// TIA Portal V20 program export: 15 tag tables, 7 data types, 9 data blocks, 10 code blocks (in call order from the OBs), 5 instance data blocks

VAR_GLOBAL   // PLC tag table "COGNEX_ETIKETA"
   "COG_ETIKETA_COG_ETIKETA_is3800-TriggerEnable" AT %Q2.0 : Bool;
   "COG_ETIKETA_COG_ETIKETA_is3800-Trigger" AT %Q2.1 : Bool;
   "COG_ETIKETA_is3800-ClearExposureComplete" AT %Q2.2 : Bool;
   "COG_ETIKETA_is3800-Set Offline" AT %Q2.7 : Bool;
   "COG_ETIKETA_is3800-TriggerReady" AT %I2.0 : Bool;
   "COG_ETIKETA_is3800-TriggerAck" AT %I2.1 : Bool;
   "COG_ETIKETA_is3800-ExposureComplete" AT %I2.2 : Bool;
   "COG_ETIKETA_is3800-AcquCOG_ETIKETA_isitionError" AT %I2.3 : Bool;
   "COG_ETIKETA_is3800-Offline Reason" AT %I2.4 : Bool;
   "COG_ETIKETA_is3800-Offline Reason(1)" AT %I2.5 : Bool;
   "COG_ETIKETA_is3800-Offline Reason(2)" AT %I2.6 : Bool;
   "COG_ETIKETA_is3800-Online" AT %I2.7 : Bool;
   "COG_ETIKETA_is3800-AcquCOG_ETIKETA_isitionID" AT %IW4 : Int;
   "COG_ETIKETA_is3800-BufferResultsEnable" AT %Q3.0 : Bool;
   "COG_ETIKETA_is3800-InspectionResultsAck" AT %Q3.1 : Bool;
   "COG_ETIKETA_is3800-SetUserData" AT %Q3.2 : Bool;
   "COG_ETIKETA_is3800-ExecuteCommand/JobLoad" AT %Q3.3 : Bool;
   "COG_ETIKETA_is3800-ClearError" AT %Q3.7 : Bool;
   "COG_ETIKETA_is3800-Reserved" AT %I10.0 : Bool;
   "COG_ETIKETA_is3800-InspectionCompleted" AT %I10.1 : Bool;
   "COG_ETIKETA_is3800-ResultsBufferOverrun" AT %I10.2 : Bool;
   "COG_ETIKETA_is3800-ResultsValid" AT %I10.3 : Bool;
   "COG_ETIKETA_is3800-CommandExecuting" AT %I10.4 : Bool;
   "COG_ETIKETA_is3800-CommandCompleted" AT %I10.5 : Bool;
   "COG_ETIKETA_is3800-CommandFailed" AT %I10.6 : Bool;
   "COG_ETIKETA_is3800-SetUserDataAck" AT %I10.7 : Bool;
   "COG_ETIKETA_is3800-ResultsPassed (Job)" AT %I11.0 : Bool;
   "COG_ETIKETA_is3800-SystemValidated" AT %I11.1 : Bool;
   "COG_ETIKETA_is3800-Error" AT %I11.7 : Bool;
   "COG_ETIKETA_is3800-ErrorCode" AT %IW12 : Word;
   "COG_ETIKETA_is3800-CommandID" AT %QW64 : Word;
   "COG_ETIKETA_is3800-Current Job ID" AT %IW68 : Word;
   "COG_ETIKETA_is3800-CommandResultCode" AT %IW70 : Word;
   "COG_ETIKETA_is3800-ExternalEvent[0]" AT %Q4.0 : Bool;
   "COG_ETIKETA_is3800-ExternalEvent[1]" AT %Q4.1 : Bool;
   "COG_ETIKETA_is3800-ExternalEvent[2]" AT %Q4.2 : Bool;
   "COG_ETIKETA_is3800-ExternalEvent[3]" AT %Q4.3 : Bool;
   "COG_ETIKETA_is3800-ExternalEvent[4]" AT %Q4.4 : Bool;
   "COG_ETIKETA_is3800-ExternalEvent[5]" AT %Q4.5 : Bool;
   "COG_ETIKETA_is3800-ExternalEvent[6]" AT %Q4.6 : Bool;
   "COG_ETIKETA_is3800-ExternalEvent[7]" AT %Q4.7 : Bool;
   "COG_ETIKETA_is3800-ExternalEventAck[0]" AT %I6.0 : Bool;
   "COG_ETIKETA_is3800-ExternalEventAck[1]" AT %I6.1 : Bool;
   "COG_ETIKETA_is3800-ExternalEventAck[2]" AT %I6.2 : Bool;
   "COG_ETIKETA_is3800-ExternalEventAck[3]" AT %I6.3 : Bool;
   "COG_ETIKETA_is3800-ExternalEventAck[4]" AT %I6.4 : Bool;
   "COG_ETIKETA_is3800-ExternalEventAck[5]" AT %I6.5 : Bool;
   "COG_ETIKETA_is3800-ExternalEventAck[6]" AT %I6.6 : Bool;
   "COG_ETIKETA_is3800-ExternalEventAck[7]" AT %I6.7 : Bool;
   "COG_ETIKETA_is3800-UserData[0]" AT %QB66 : Byte;
   "COG_ETIKETA_is3800-UserData[1]" AT %QB67 : Byte;
   "COG_ETIKETA_is3800-UserData[2]" AT %QB68 : Byte;
   "COG_ETIKETA_is3800-UserData[3]" AT %QB69 : Byte;
   "COG_ETIKETA_is3800-UserData[4]" AT %QB70 : Byte;
   "COG_ETIKETA_is3800-UserData[5]" AT %QB71 : Byte;
   "COG_ETIKETA_is3800-UserData[6]" AT %QB72 : Byte;
   "COG_ETIKETA_is3800-UserData[7]" AT %QB73 : Byte;
   "COG_ETIKETA_is3800-UserData[8]" AT %QB74 : Byte;
   "COG_ETIKETA_is3800-UserData[9]" AT %QB75 : Byte;
   "COG_ETIKETA_is3800-UserData[10]" AT %QB76 : Byte;
   "COG_ETIKETA_is3800-UserData[11]" AT %QB77 : Byte;
   "COG_ETIKETA_is3800-UserData[12]" AT %QB78 : Byte;
   "COG_ETIKETA_is3800-UserData[13]" AT %QB79 : Byte;
   "COG_ETIKETA_is3800-UserData[14]" AT %QB80 : Byte;
   "COG_ETIKETA_is3800-UserData[15]" AT %QB81 : Byte;
   "COG_ETIKETA_is3800-InspectionID" AT %IW72 : Word;
   "COG_ETIKETA_is3800-InspectionResultsCode" AT %IW74 : Int;
   "COG_ETIKETA_is3800-InspectionResults_0" AT %IB76 : Byte;
   "COG_ETIKETA_is3800-InspectionResults_1" AT %IB77 : Byte;
   "COG_ETIKETA_is3800-InspectionResults_2" AT %IB78 : Byte;
   "COG_ETIKETA_is3800-InspectionResults_3" AT %IB79 : Byte;
   "COG_ETIKETA_is3800-InspectionResults_4" AT %IB80 : Byte;
   "COG_ETIKETA_is3800-InspectionResults_5" AT %IB81 : Byte;
   "COG_ETIKETA_is3800-InspectionResults_6" AT %IB82 : Byte;
   "COG_ETIKETA_is3800-InspectionResults_7" AT %IB83 : Byte;
   "COG_ETIKETA_is3800-InspectionResults_8" AT %IB84 : Byte;
   "COG_ETIKETA_is3800-InspectionResults_9" AT %IB85 : Byte;
   "COG_ETIKETA_is3800-InspectionResults_10" AT %IB86 : Byte;
   "COG_ETIKETA_is3800-InspectionResults_11" AT %IB87 : Byte;
   "COG_ETIKETA_is3800-InspectionResults_12" AT %IB88 : Byte;
   "COG_ETIKETA_is3800-InspectionResults_13" AT %IB89 : Byte;
   "COG_ETIKETA_is3800-InspectionResults_14" AT %IB90 : Byte;
   "COG_ETIKETA_is3800-InspectionResults_15" AT %IB91 : Byte;
   "COG_ETIKETA_is3800-InspectionResults_16" AT %IB92 : Byte;
   "COG_ETIKETA_is3800-InspectionResults_17" AT %IB93 : Byte;
   "COG_ETIKETA_is3800-InspectionResults_18" AT %IB94 : Byte;
   "COG_ETIKETA_is3800-InspectionResults_19" AT %IB95 : Byte;
   "COG_ETIKETA_is3800-InspectionResults_20" AT %IB96 : Byte;
   "COG_ETIKETA_is3800-InspectionResults_21" AT %IB97 : Byte;
   "COG_ETIKETA_is3800-InspectionResults_22" AT %IB98 : Byte;
   "COG_ETIKETA_is3800-InspectionResults_23" AT %IB99 : Byte;
   "COG_ETIKETA_is3800-InspectionResults_24" AT %IB100 : Byte;
   "COG_ETIKETA_is3800-InspectionResults_25" AT %IB101 : Byte;
   "COG_ETIKETA_is3800-InspectionResults_26" AT %IB102 : Byte;
   "COG_ETIKETA_is3800-InspectionResults_27" AT %IB103 : Byte;
   "COG_ETIKETA_is3800-InspectionResults_28" AT %IB104 : Byte;
   "COG_ETIKETA_is3800-InspectionResults_29" AT %IB105 : Byte;
   "COG_ETIKETA_is3800-InspectionResults_30" AT %IB106 : Byte;
   "COG_ETIKETA_is3800-InspectionResults_31" AT %IB107 : Byte;
   "COG_ETIKETA_is3800-InspectionResults_32" AT %IB108 : Byte;
   "COG_ETIKETA_is3800-InspectionResults_33" AT %IB109 : Byte;
   "COG_ETIKETA_is3800-InspectionResults_34" AT %IB110 : Byte;
   "COG_ETIKETA_is3800-InspectionResults_35" AT %IB111 : Byte;
   "COG_ETIKETA_is3800-InspectionResults_36" AT %IB112 : Byte;
   "COG_ETIKETA_is3800-InspectionResults_37" AT %IB113 : Byte;
   "COG_ETIKETA_is3800-InspectionResults_38" AT %IB114 : Byte;
   "COG_ETIKETA_is3800-InspectionResults_39" AT %IB115 : Byte;
   "COG_ETIKETA_is3800-InspectionResults_40" AT %IB116 : Byte;
   "COG_ETIKETA_is3800-InspectionResults_41" AT %IB117 : Byte;
   "COG_ETIKETA_is3800-InspectionResults_42" AT %IB118 : Byte;
   "COG_ETIKETA_is3800-InspectionResults_43" AT %IB119 : Byte;
   "COG_ETIKETA_is3800-InspectionResults_44" AT %IB120 : Byte;
   "COG_ETIKETA_is3800-InspectionResults_45" AT %IB121 : Byte;
   "COG_ETIKETA_is3800-InspectionResults_46" AT %IB122 : Byte;
   "COG_ETIKETA_is3800-InspectionResults_47" AT %IB123 : Byte;
   "COG_ETIKETA_is3800-InspectionResults_48" AT %IB124 : Byte;
   "COG_ETIKETA_is3800-InspectionResults_49" AT %IB125 : Byte;
   "COG_ETIKETA_is3800-InspectionResults_50" AT %IB126 : Byte;
   "COG_ETIKETA_is3800-InspectionResults_51" AT %IB127 : Byte;
   "COG_ETIKETA_is3800-InspectionResults_52" AT %IB128 : Byte;
   "COG_ETIKETA_is3800-InspectionResults_53" AT %IB129 : Byte;
   "COG_ETIKETA_is3800-InspectionResults_54" AT %IB130 : Byte;
   "COG_ETIKETA_is3800-InspectionResults_55" AT %IB131 : Byte;
   "COG_ETIKETA_is3800-InspectionResults_56" AT %IB132 : Byte;
   "COG_ETIKETA_is3800-InspectionResults_57" AT %IB133 : Byte;
   "COG_ETIKETA_is3800-InspectionResults_58" AT %IB134 : Byte;
   "COG_ETIKETA_is3800-InspectionResults_59" AT %IB135 : Byte;
   "COG_ETIKETA_is3800-InspectionResults_60" AT %IB136 : Byte;
   "COG_ETIKETA_is3800-InspectionResults_61" AT %IB137 : Byte;
   "COG_ETIKETA_is3800-InspectionResults_62" AT %IB138 : Byte;
   "COG_ETIKETA_is3800-InspectionResults_63" AT %IB139 : Byte;
   "COG_ETIKETA_is3800-InspectionResults_64" AT %IB140 : Byte;
   "COG_ETIKETA_is3800-InspectionResults_65" AT %IB141 : Byte;
   "COG_ETIKETA_is3800-InspectionResults_66" AT %IB142 : Byte;
   "COG_ETIKETA_is3800-InspectionResults_67" AT %IB143 : Byte;
   "COG_ETIKETA_is3800-InspectionResults_68" AT %IB144 : Byte;
   "COG_ETIKETA_is3800-InspectionResults_69" AT %IB145 : Byte;
   "COG_ETIKETA_is3800-InspectionResults_70" AT %IB146 : Byte;
   "COG_ETIKETA_is3800-InspectionResults_71" AT %IB147 : Byte;
   "COG_ETIKETA_is3800-InspectionResults_72" AT %IB148 : Byte;
   "COG_ETIKETA_is3800-InspectionResults_73" AT %IB149 : Byte;
   "COG_ETIKETA_is3800-InspectionResults_74" AT %IB150 : Byte;
   "COG_ETIKETA_is3800-InspectionResults_75" AT %IB151 : Byte;
   "COG_ETIKETA_is3800-InspectionResults_76" AT %IB152 : Byte;
   "COG_ETIKETA_is3800-InspectionResults_77" AT %IB153 : Byte;
   "COG_ETIKETA_is3800-InspectionResults_78" AT %IB154 : Byte;
   "COG_ETIKETA_is3800-InspectionResults_79" AT %IB155 : Byte;
   "COG_ETIKETA_is3800-InspectionResults_80" AT %IB156 : Byte;
   "COG_ETIKETA_is3800-InspectionResults_81" AT %IB157 : Byte;
   "COG_ETIKETA_is3800-InspectionResults_82" AT %IB158 : Byte;
   "COG_ETIKETA_is3800-InspectionResults_83" AT %IB159 : Byte;
   "COG_ETIKETA_is3800-InspectionResults_84" AT %IB160 : Byte;
   "COG_ETIKETA_is3800-InspectionResults_85" AT %IB164 : Byte;
   "COG_ETIKETA_is3800-InspectionResults_86" AT %IB165 : Byte;
   "COG_ETIKETA_is3800-InspectionResults_87" AT %IB166 : Byte;
   "COG_ETIKETA_is3800-InspectionResults_88" AT %IB167 : Byte;
   "COG_ETIKETA_is3800-InspectionResults_89" AT %IB168 : Byte;
   "COG_ETIKETA_is3800-InspectionResults_90" AT %IB169 : Byte;
   "COG_ETIKETA_is3800-InspectionResults_91" AT %IB170 : Byte;
   "COG_ETIKETA_is3800-InspectionResults_92" AT %IB171 : Byte;
   "COG_ETIKETA_is3800-InspectionResults_93" AT %IB172 : Byte;
   "COG_ETIKETA_is3800-InspectionResults_94" AT %IB173 : Byte;
   "COG_ETIKETA_is3800-InspectionResults_95" AT %IB174 : Byte;
   "COG_ETIKETA_is3800-InspectionResults_96" AT %IB175 : Byte;
   "COG_ETIKETA_is3800-InspectionResults_97" AT %IB176 : Byte;
   "COG_ETIKETA_is3800-InspectionResults_98" AT %IB177 : Byte;
   "COG_ETIKETA_is3800-InspectionResults_99" AT %IB178 : Byte;
   "COG_ETIKETA_is3800-InspectionResults_100" AT %IB179 : Byte;
END_VAR

VAR_GLOBAL   // PLC tag table "COGNEX_FOLIE_L"
   "COG_FOLIE_L_COG_FOLIE_L_is3800-TriggerEnable" AT %Q5.0 : Bool;
   "COG_FOLIE_L_is3800-Trigger" AT %Q5.1 : Bool;
   "COG_FOLIE_L_is3800-ClearExposureComplete" AT %Q5.2 : Bool;
   "COG_FOLIE_L_is3800-Set Offline" AT %Q5.7 : Bool;
   "COG_FOLIE_L_is3800-TriggerReady" AT %I14.0 : Bool;
   "COG_FOLIE_L_is3800-TriggerAck" AT %I14.1 : Bool;
   "COG_FOLIE_L_is3800-ExposureComplete" AT %I14.2 : Bool;
   "COG_FOLIE_L_is3800-AcquCOG_FOLIE_L_isitionError" AT %I14.3 : Bool;
   "COG_FOLIE_L_is3800-Offline Reason" AT %I14.4 : Bool;
   "COG_FOLIE_L_is3800-Offline Reason(1)" AT %I14.5 : Bool;
   "COG_FOLIE_L_is3800-Offline Reason(2)" AT %I14.6 : Bool;
   "COG_FOLIE_L_is3800-Online" AT %I14.7 : Bool;
   "COG_FOLIE_L_is3800-AcquCOG_FOLIE_L_isitionID" AT %IW16 : Int;
   "COG_FOLIE_L_is3800-BufferResultsEnable" AT %Q6.0 : Bool;
   "COG_FOLIE_L_is3800-InspectionResultsAck" AT %Q6.1 : Bool;
   "COG_FOLIE_L_is3800-SetUserData" AT %Q6.2 : Bool;
   "COG_FOLIE_L_is3800-ExecuteCommand/JobLoad" AT %Q6.3 : Bool;
   "COG_FOLIE_L_is3800-ClearError" AT %Q6.7 : Bool;
   "COG_FOLIE_L_is3800-Reserved" AT %I18.0 : Bool;
   "COG_FOLIE_L_is3800-InspectionCompleted" AT %I18.1 : Bool;
   "COG_FOLIE_L_is3800-ResultsBufferOverrun" AT %I18.2 : Bool;
   "COG_FOLIE_L_is3800-ResultsValid" AT %I18.3 : Bool;
   "COG_FOLIE_L_is3800-CommandExecuting" AT %I18.4 : Bool;
   "COG_FOLIE_L_is3800-CommandCompleted" AT %I18.5 : Bool;
   "COG_FOLIE_L_is3800-CommandFailed" AT %I18.6 : Bool;
   "COG_FOLIE_L_is3800-SetUserDataAck" AT %I18.7 : Bool;
   "COG_FOLIE_L_is3800-ResultsPassed (Job)" AT %I19.0 : Bool;
   "COG_FOLIE_L_is3800-SystemValidated" AT %I19.1 : Bool;
   "COG_FOLIE_L_is3800-Error" AT %I19.7 : Bool;
   "COG_FOLIE_L_is3800-ErrorCode" AT %IW20 : Word;
   "COG_FOLIE_L_is3800-CommandID" AT %QW130 : Word;
   "COG_FOLIE_L_is3800-Current Job ID" AT %IW140 : Word;
   "COG_FOLIE_L_is3800-CommandResultCode" AT %IW142 : Word;
   "COG_FOLIE_L_is3800-ExternalEvent[0]" AT %Q7.0 : Bool;
   "COG_FOLIE_L_is3800-ExternalEvent[1]" AT %Q7.1 : Bool;
   "COG_FOLIE_L_is3800-ExternalEvent[2]" AT %Q7.2 : Bool;
   "COG_FOLIE_L_is3800-ExternalEvent[3]" AT %Q7.3 : Bool;
   "COG_FOLIE_L_is3800-ExternalEvent[4]" AT %Q7.4 : Bool;
   "COG_FOLIE_L_is3800-ExternalEvent[5]" AT %Q7.5 : Bool;
   "COG_FOLIE_L_is3800-ExternalEvent[6]" AT %Q7.6 : Bool;
   "COG_FOLIE_L_is3800-ExternalEvent[7]" AT %Q7.7 : Bool;
   "COG_FOLIE_L_is3800-ExternalEventAck[0]" AT %I7.0 : Bool;
   "COG_FOLIE_L_is3800-ExternalEventAck[1]" AT %I7.1 : Bool;
   "COG_FOLIE_L_is3800-ExternalEventAck[2]" AT %I7.2 : Bool;
   "COG_FOLIE_L_is3800-ExternalEventAck[3]" AT %I7.3 : Bool;
   "COG_FOLIE_L_is3800-ExternalEventAck[4]" AT %I7.4 : Bool;
   "COG_FOLIE_L_is3800-ExternalEventAck[5]" AT %I7.5 : Bool;
   "COG_FOLIE_L_is3800-ExternalEventAck[6]" AT %I7.6 : Bool;
   "COG_FOLIE_L_is3800-ExternalEventAck[7]" AT %I7.7 : Bool;
   "COG_FOLIE_L_is3800-UserData[0]" AT %QB132 : Byte;
   "COG_FOLIE_L_is3800-UserData[1]" AT %QB133 : Byte;
   "COG_FOLIE_L_is3800-UserData[2]" AT %QB134 : Byte;
   "COG_FOLIE_L_is3800-UserData[3]" AT %QB135 : Byte;
   "COG_FOLIE_L_is3800-UserData[4]" AT %QB136 : Byte;
   "COG_FOLIE_L_is3800-UserData[5]" AT %QB137 : Byte;
   "COG_FOLIE_L_is3800-UserData[6]" AT %QB138 : Byte;
   "COG_FOLIE_L_is3800-UserData[7]" AT %QB139 : Byte;
   "COG_FOLIE_L_is3800-UserData[8]" AT %QB140 : Byte;
   "COG_FOLIE_L_is3800-UserData[9]" AT %QB141 : Byte;
   "COG_FOLIE_L_is3800-UserData[10]" AT %QB142 : Byte;
   "COG_FOLIE_L_is3800-UserData[11]" AT %QB143 : Byte;
   "COG_FOLIE_L_is3800-UserData[12]" AT %QB144 : Byte;
   "COG_FOLIE_L_is3800-UserData[13]" AT %QB145 : Byte;
   "COG_FOLIE_L_is3800-UserData[14]" AT %QB146 : Byte;
   "COG_FOLIE_L_is3800-UserData[15]" AT %QB147 : Byte;
   "COG_FOLIE_L_is3800-InspectionID" AT %IW144 : Word;
   "COG_FOLIE_L_is3800-InspectionResultsCode" AT %IW146 : Int;
   "COG_FOLIE_L_is3800-InspectionResults[0]" AT %IB148 : Byte;
   "COG_FOLIE_L_is3800-InspectionResults[1]" AT %IB149 : Byte;
   "COG_FOLIE_L_is3800-InspectionResults[2]" AT %IB150 : Byte;
   "COG_FOLIE_L_is3800-InspectionResults[3]" AT %IB151 : Byte;
   "COG_FOLIE_L_is3800-InspectionResults[4]" AT %IB152 : Byte;
   "COG_FOLIE_L_is3800-InspectionResults[5]" AT %IB153 : Byte;
   "COG_FOLIE_L_is3800-InspectionResults[6]" AT %IB154 : Byte;
   "COG_FOLIE_L_is3800-InspectionResults[7]" AT %IB155 : Byte;
   "COG_FOLIE_L_is3800-InspectionResults[8]" AT %IB156 : Byte;
   "COG_FOLIE_L_is3800-InspectionResults[9]" AT %IB157 : Byte;
   "COG_FOLIE_L_is3800-InspectionResults[10]" AT %IB158 : Byte;
   "COG_FOLIE_L_is3800-InspectionResults[11]" AT %IB159 : Byte;
   "COG_FOLIE_L_is3800-InspectionResults[12]" AT %IB160 : Byte;
   "COG_FOLIE_L_is3800-InspectionResults[13]" AT %IB161 : Byte;
   "COG_FOLIE_L_is3800-InspectionResults[14]" AT %IB162 : Byte;
   "COG_FOLIE_L_is3800-InspectionResults[15]" AT %IB163 : Byte;
END_VAR

VAR_GLOBAL   // PLC tag table "COGNEX_FOLIE_P"
   "COG_FOLIE_P_COG_FOLIE_P_is3800-TriggerEnable" AT %Q10.0 : Bool;
   "COG_FOLIE_P_is3800-Trigger" AT %Q10.1 : Bool;
   "COG_FOLIE_P_is3800-ClearExposureComplete" AT %Q10.2 : Bool;
   "COG_FOLIE_P_is3800-Set Offline" AT %Q10.7 : Bool;
   "COG_FOLIE_P_is3800-TriggerReady" AT %I22.0 : Bool;
   "COG_FOLIE_P_is3800-TriggerAck" AT %I22.1 : Bool;
   "COG_FOLIE_P_is3800-ExposureComplete" AT %I22.2 : Bool;
   "COG_FOLIE_P_is3800-AcquCOG_FOLIE_P_isitionError" AT %I22.3 : Bool;
   "COG_FOLIE_P_is3800-Offline Reason" AT %I22.4 : Bool;
   "COG_FOLIE_P_is3800-Offline Reason(1)" AT %I22.5 : Bool;
   "COG_FOLIE_P_is3800-Offline Reason(2)" AT %I22.6 : Bool;
   "COG_FOLIE_P_is3800-Online" AT %I22.7 : Bool;
   "COG_FOLIE_P_is3800-AcquCOG_FOLIE_P_isitionID" AT %IW24 : Int;
   "COG_FOLIE_P_is3800-BufferResultsEnable" AT %Q11.0 : Bool;
   "COG_FOLIE_P_is3800-InspectionResultsAck" AT %Q11.1 : Bool;
   "COG_FOLIE_P_is3800-SetUserData" AT %Q11.2 : Bool;
   "COG_FOLIE_P_is3800-ExecuteCommand/JobLoad" AT %Q11.3 : Bool;
   "COG_FOLIE_P_is3800-ClearError" AT %Q11.7 : Bool;
   "COG_FOLIE_P_is3800-Reserved" AT %I26.0 : Bool;
   "COG_FOLIE_P_is3800-InspectionCompleted" AT %I26.1 : Bool;
   "COG_FOLIE_P_is3800-ResultsBufferOverrun" AT %I26.2 : Bool;
   "COG_FOLIE_P_is3800-ResultsValid" AT %I26.3 : Bool;
   "COG_FOLIE_P_is3800-CommandExecuting" AT %I26.4 : Bool;
   "COG_FOLIE_P_is3800-CommandCompleted" AT %I26.5 : Bool;
   "COG_FOLIE_P_is3800-CommandFailed" AT %I26.6 : Bool;
   "COG_FOLIE_P_is3800-SetUserDataAck" AT %I26.7 : Bool;
   "COG_FOLIE_P_is3800-ResultsPassed (Job)" AT %I27.0 : Bool;
   "COG_FOLIE_P_is3800-SystemValidated" AT %I27.1 : Bool;
   "COG_FOLIE_P_is3800-Error" AT %I27.7 : Bool;
   "COG_FOLIE_P_is3800-ErrorCode" AT %IW28 : Word;
   "COG_FOLIE_P_is3800-CommandID" AT %QW196 : Word;
   "COG_FOLIE_P_is3800-Current Job ID" AT %IW212 : Word;
   "COG_FOLIE_P_is3800-CommandResultCode" AT %IW214 : Word;
   "COG_FOLIE_P_is3800-ExternalEvent[0]" AT %Q12.0 : Bool;
   "COG_FOLIE_P_is3800-ExternalEvent[1]" AT %Q12.1 : Bool;
   "COG_FOLIE_P_is3800-ExternalEvent[2]" AT %Q12.2 : Bool;
   "COG_FOLIE_P_is3800-ExternalEvent[3]" AT %Q12.3 : Bool;
   "COG_FOLIE_P_is3800-ExternalEvent[4]" AT %Q12.4 : Bool;
   "COG_FOLIE_P_is3800-ExternalEvent[5]" AT %Q12.5 : Bool;
   "COG_FOLIE_P_is3800-ExternalEvent[6]" AT %Q12.6 : Bool;
   "COG_FOLIE_P_is3800-ExternalEvent[7]" AT %Q12.7 : Bool;
   "COG_FOLIE_P_is3800-ExternalEventAck[0]" AT %I30.0 : Bool;
   "COG_FOLIE_P_is3800-ExternalEventAck[1]" AT %I30.1 : Bool;
   "COG_FOLIE_P_is3800-ExternalEventAck[2]" AT %I30.2 : Bool;
   "COG_FOLIE_P_is3800-ExternalEventAck[3]" AT %I30.3 : Bool;
   "COG_FOLIE_P_is3800-ExternalEventAck[4]" AT %I30.4 : Bool;
   "COG_FOLIE_P_is3800-ExternalEventAck[5]" AT %I30.5 : Bool;
   "COG_FOLIE_P_is3800-ExternalEventAck[6]" AT %I30.6 : Bool;
   "COG_FOLIE_P_is3800-ExternalEventAck[7]" AT %I30.7 : Bool;
   "COG_FOLIE_P_is3800-UserData[0]" AT %QB198 : Byte;
   "COG_FOLIE_P_is3800-UserData[1]" AT %QB199 : Byte;
   "COG_FOLIE_P_is3800-UserData[2]" AT %QB200 : Byte;
   "COG_FOLIE_P_is3800-UserData[3]" AT %QB201 : Byte;
   "COG_FOLIE_P_is3800-UserData[4]" AT %QB202 : Byte;
   "COG_FOLIE_P_is3800-UserData[5]" AT %QB203 : Byte;
   "COG_FOLIE_P_is3800-UserData[6]" AT %QB204 : Byte;
   "COG_FOLIE_P_is3800-UserData[7]" AT %QB205 : Byte;
   "COG_FOLIE_P_is3800-UserData[8]" AT %QB206 : Byte;
   "COG_FOLIE_P_is3800-UserData[9]" AT %QB207 : Byte;
   "COG_FOLIE_P_is3800-UserData[10]" AT %QB208 : Byte;
   "COG_FOLIE_P_is3800-UserData[11]" AT %QB209 : Byte;
   "COG_FOLIE_P_is3800-UserData[12]" AT %QB210 : Byte;
   "COG_FOLIE_P_is3800-UserData[13]" AT %QB211 : Byte;
   "COG_FOLIE_P_is3800-UserData[14]" AT %QB212 : Byte;
   "COG_FOLIE_P_is3800-UserData[15]" AT %QB213 : Byte;
   "COG_FOLIE_P_is3800-InspectionID" AT %IW216 : Word;
   "COG_FOLIE_P_is3800-InspectionResultsCode" AT %IW218 : Int;
   "COG_FOLIE_P_is3800-InspectionResults[0]" AT %IB220 : Byte;
   "COG_FOLIE_P_is3800-InspectionResults[1]" AT %IB221 : Byte;
   "COG_FOLIE_P_is3800-InspectionResults[2]" AT %IB222 : Byte;
   "COG_FOLIE_P_is3800-InspectionResults[3]" AT %IB223 : Byte;
   "COG_FOLIE_P_is3800-InspectionResults[4]" AT %IB224 : Byte;
   "COG_FOLIE_P_is3800-InspectionResults[5]" AT %IB225 : Byte;
   "COG_FOLIE_P_is3800-InspectionResults[6]" AT %IB226 : Byte;
   "COG_FOLIE_P_is3800-InspectionResults[7]" AT %IB227 : Byte;
   "COG_FOLIE_P_is3800-InspectionResults[8]" AT %IB228 : Byte;
   "COG_FOLIE_P_is3800-InspectionResults[9]" AT %IB229 : Byte;
   "COG_FOLIE_P_is3800-InspectionResults[10]" AT %IB230 : Byte;
   "COG_FOLIE_P_is3800-InspectionResults[11]" AT %IB231 : Byte;
   "COG_FOLIE_P_is3800-InspectionResults[12]" AT %IB232 : Byte;
   "COG_FOLIE_P_is3800-InspectionResults[13]" AT %IB233 : Byte;
   "COG_FOLIE_P_is3800-InspectionResults[14]" AT %IB234 : Byte;
   "COG_FOLIE_P_is3800-InspectionResults[15]" AT %IB235 : Byte;
END_VAR

VAR_GLOBAL   // PLC tag table "Default tag table"
   RESERVE_AI_1 AT %IW66 : Int;
   "System_Byte(1)" AT %MB1 : Byte;
   reset_hsc AT %M2.7 : Bool;
END_VAR

VAR_GLOBAL   // PLC tag table "PLC-A3-AI"
   RESERVE_AI AT %IW64 : Int;
END_VAR

VAR_GLOBAL   // PLC tag table "PLC-A3-DI"
   "ENCODER_L+" AT %I0.0 : Bool;   // JEDEN ENCODER DVA KANÁLY NAASTAVENÍ NA HSPEED COUNTER
   "ENCODER_L-" AT %I0.1 : Bool;   // JEDEN ENCODER DVA KANÁLY NAASTAVENÍ NA HSPEED COUNTER
   ENCODER AT %I0.2 : Bool;
   "ENCODER(1)" AT %I0.3 : Bool;
   "ENCODER(2)" AT %I0.4 : Bool;
   RESERVE_DI AT %I0.5 : Bool;   // s1 najezd
   RESERVE_DI_1 AT %I0.6 : Bool;   // s2 foceni
   RESERVE_DI_2 AT %I0.7 : Bool;   // s3 konec budky
   RESERVE_DI_3 AT %I1.0 : Bool;   // s4 vyrazovač
   RESERVE_DI_4 AT %I1.1 : Bool;   // s5 valec pozice home
   RESERVE_DI_5 AT %I1.2 : Bool;
   RESERVE_DI_6 AT %I1.3 : Bool;
   RESERVE_DI_7 AT %I1.4 : Bool;
   RESERVE_DI_8 AT %I1.5 : Bool;
END_VAR

VAR_GLOBAL   // PLC tag table "PLC-A3-DQ"
   "-KA1" AT %Q0.0 : Bool;   // OSVĚTLENÍ FOLIE
   "-KA2" AT %Q0.1 : Bool;   // OSVĚTLENÍ FOLIE
   "-KA3" AT %Q0.2 : Bool;   // OSVĚTLENÍ FOLIE
   "-KA4" AT %Q0.3 : Bool;   // OSVĚTLENÍ ETIKETA
   "-KA5" AT %Q0.4 : Bool;   // OSVĚTLENÍ ETIKETA
   "-KA18" AT %Q0.5 : Bool;   // MAJÁK_žlutá
   "-KA19" AT %Q0.6 : Bool;   // MAJÁK_červená
   "-KA20" AT %Q0.7 : Bool;   // MAJÁK_zelena
   "-KA21" AT %Q1.0 : Bool;   // HOUKAČKA
   RESERVE_DQ AT %Q1.1 : Bool;
END_VAR

VAR_GLOBAL   // PLC tag table "PLC-A4-DI"
   "-KA6" AT %I8.0 : Bool;
   "-KA7" AT %I8.1 : Bool;
   "-KA8" AT %I8.2 : Bool;
   "-KA9" AT %I8.3 : Bool;
   "-KA10" AT %I8.4 : Bool;
   "-KA11" AT %I8.5 : Bool;
   RESERVE_DI_9 AT %I8.6 : Bool;
   RESERVE_DI_10 AT %I8.7 : Bool;
   RESERVE_DI_11 AT %I9.0 : Bool;   // dveře L kanál A
   RESERVE_DI_12 AT %I9.1 : Bool;   // dveře L kanál B
   RESERVE_DI_13 AT %I9.2 : Bool;   // dveře P kanál A
   RESERVE_DI_14 AT %I9.3 : Bool;   // Dveře P kanál B
   RESERVE_DI_15 AT %I9.4 : Bool;
   RESERVE_DI_16 AT %I9.5 : Bool;
   RESERVE_DI_17 AT %I9.6 : Bool;
   RESERVE_DI_18 AT %I9.7 : Bool;
END_VAR

VAR_GLOBAL   // PLC tag table "PLC-A4-DQ"
   "-KA12" AT %Q8.0 : Bool;
   "-KA13" AT %Q8.1 : Bool;
   "-KA14" AT %Q8.2 : Bool;
   "-KA15" AT %Q8.3 : Bool;
   "-KA16" AT %Q8.4 : Bool;
   "-KA17" AT %Q8.5 : Bool;
   RESERVE_DQ_ AT %Q8.6 : Bool;
   RESERVE_DQ_1 AT %Q8.7 : Bool;
   RESERVE_DQ_2 AT %Q9.0 : Bool;   // vyrazovac
   RESERVE_DQ_3 AT %Q9.1 : Bool;
   RESERVE_DQ_4 AT %Q9.2 : Bool;
   RESERVE_DQ_5 AT %Q9.3 : Bool;
   RESERVE_DQ_6 AT %Q9.4 : Bool;
   RESERVE_DQ_7 AT %Q9.5 : Bool;
   RESERVE_DQ_8 AT %Q9.6 : Bool;
   RESERVE_DQ_9 AT %Q9.7 : Bool;
END_VAR

VAR_GLOBAL   // PLC tag table "memor"
   HSC_1 AT %ID1000 : DWord;
   PAMET_TEST AT %MD16 : DInt;
   ret_val_move_blk AT %MW20 : Int;
   i AT %MW22 : Int;
   "i(1)" AT %MW24 : Int;
END_VAR

VAR_GLOBAL   // PLC tag table "standard"
   SIMULACE AT %M2.0 : Bool;
   LOG_0 AT %M2.1 : Bool;
   LOG_1 AT %M2.2 : Bool;
   SMAZ_ME_0 AT %M2.3 : Bool;
   SMAZ_ME_1 AT %M2.4 : Bool;
   AUTOMAT AT %M2.5 : Bool;
   MANUAL AT %M2.6 : Bool;
   INICIALIZACE_OK AT %M3.3 : Bool;
   INICIALIZACE AT %M3.4 : Bool;
   INICIALIZACE_RUN AT %M3.5 : Bool;
   LINE_READY_START AT %M3.6 : Bool;
   alrm_global AT %M3.2 : Bool;
   wrong_global AT %M3.7 : Bool;
   alrm_op_0 AT %M4.0 : Bool;
   wrong_op_0 AT %M4.1 : Bool;
   alrm_op_1 AT %M4.2 : Bool;
   wrong_op_1 AT %M4.3 : Bool;
   I_i AT %MW6 : Int;
   "I_i(1)" AT %MW8 : Int;
   adresace AT %MW12 : Int;
   byte_smazat AT %MB5 : Byte;
   inicializace_block AT %M4.4 : Bool;
   s2_hsc_hrana AT %M4.5 : Bool;
   hodnota_volitelna AT %MB14 : Byte;
   Clock_Byte AT %MB0 : Byte;
   Clock_10Hz AT %M0.0 : Bool;
   Clock_5Hz AT %M0.1 : Bool;
   "Clock_2.5Hz" AT %M0.2 : Bool;
   Clock_2Hz AT %M0.3 : Bool;
   "Clock_1.25Hz" AT %M0.4 : Bool;
   Clock_1Hz AT %M0.5 : Bool;
   "Clock_0.625Hz" AT %M0.6 : Bool;
   "Clock_0.5Hz" AT %M0.7 : Bool;
   System_Byte AT %MB1 : Byte;
   FirstScan AT %M1.0 : Bool;
   DiagStatusUpdate AT %M1.1 : Bool;
   AlwaysTRUE AT %M1.2 : Bool;
   AlwaysFALSE AT %M1.3 : Bool;
   INICIALIZACE_REPEAT AT %M4.6 : Bool;
   AUT_MAN_HMI AT %M4.7 : Bool;   // POUŽÍVÁNO PRO PANELOUVOU VOLBU
   volny_pristup_2 AT %M10.0 : Bool;
   alrm_op_2 AT %M11.3 : Bool;
   wrong_op_2 AT %M11.4 : Bool;
   alrm_op_3 AT %M11.5 : Bool;
   wrong_op_3 AT %M11.6 : Bool;
   alrm_op_4 AT %M11.7 : Bool;
   wrong_op_4 AT %M15.0 : Bool;
   alrm_op_5 AT %M15.1 : Bool;
   wrong_op_5 AT %M15.2 : Bool;
   citac AT %M15.4 : Bool;
END_VAR

VAR_GLOBAL   // PLC tag table "LASER_IN_datalogic"
   LASER_OFF AT %I400.0 : Bool;
   LASER_WARM_UP AT %I400.1 : Bool;
   LASER_WAIT_FOR_START AT %I400.2 : Bool;
   LASER_STANDBY AT %I400.3 : Bool;
   LASER_STANDBY_SHUTTER_CLOSED AT %I400.4 : Bool;
   LASER_READY AT %I400.5 : Bool;
   LASER_EMISSION AT %I400.6 : Bool;
   LASER_BUSSY_SHUTTER_CLOSED AT %I401.0 : Bool;
   LASER_WARNING AT %I401.1 : Bool;
   LASER_ERROR AT %I401.2 : Bool;
   COMMAND_EXECUTING AT %I402.0 : Bool;
   COMMAND_ERROR AT %I402.1 : Bool;
   PROTOCOL_ERROR AT %I402.2 : Bool;
   PROTOCOL_BOOT_UP AT %I403.7 : Bool;
   COMMAND_ERROR_CODE AT %IB404 : Byte;
   PROTOCOL_ERROR_CODE AT %IB405 : Byte;
   RESERVE_I_6_BYTE AT %IB406 : Byte;
   RESERVE_I_7_BYTE AT %IB407 : Byte;
   RESERVE_I_8_BYTE AT %IB408 : Byte;
   RESERVE_I_9_BYTE AT %IB409 : Byte;
   START_MARKING_IN AT %I410.0 : Bool;
   STOP_SYSTEM_IN AT %I410.1 : Bool;
   GET_PNIO_PROTOCOL_VERSION_IN AT %I411.0 : Bool;
   GET_LASER_ENGINE_VERSION AT %I411.1 : Bool;
   OPEN_DOCUMENT_FROM_DEVICE AT %I412.0 : Bool;
   SAVE_DOCUMENT AT %I412.1 : Bool;
   GET_DATA_FIELD_VALUE_IN AT %I412.2 : Bool;
   SET_DATA_FIELD_VALUE_IN AT %I412.3 : Bool;
   GET_GLOBAL_COUNTER_VALUE_IN AT %I412.4 : Bool;
   SET_GLOBAL_COUNTER_VALUE_IN AT %I412.5 : Bool;
   GET_GLOBAL_STRING_VALUE_IN AT %I412.6 : Bool;
   SET_GLOBAL_STRING_VALUE_IN AT %I412.7 : Bool;
   ENABLE_DATA_FIELD_IN AT %I413.0 : Bool;
   DISABLE_DATA_FIELD_IN AT %I413.1 : Bool;
   MOVE_END_ROTATE_DOCUMENT AT %I414.0 : Bool;
   MOVE_DATA_FIELD_IN AT %I414.1 : Bool;
   RESERVE_I_15_BYTE AT %IB415 : Byte;
   RESERVE_I_16_BYTE AT %IB416 : Byte;
   RESERVE_I_17_BYTE AT %IB417 : Byte;
   MOVE_AXIS_IN AT %I418.0 : Bool;
   RESET_AXIS_IN AT %I418.1 : Bool;
   STOP_AXIS_IN AT %I418.2 : Bool;
   START_AUTOFOCUS_IN AT %I418.3 : Bool;
   STOP_AUTOFOCUS_IN AT %I418.4 : Bool;
   SET_FOCUS_DISTANCE_REFERENCE_IN AT %I418.5 : Bool;
   RESERVE_I_19_BYTE AT %IB419 : Byte;
   X_AXIS_ENABLED AT %I420.0 : Bool;
   Y_AXIS_ENABLED AT %I420.1 : Bool;
   Z_AXIS_ENABLED AT %I420.2 : Bool;
   R_AXIS_ENABLED AT %I420.3 : Bool;
   X_AXIS_HOME AT %I420.4 : Bool;
   Y_AXIS_HOME AT %I420.5 : Bool;
   Z_AXIS_HOME AT %I420.6 : Bool;
   R_AXIS_HOME AT %I420.7 : Bool;
   X_AXIS_MOVEMENT AT %I421.0 : Bool;
   Y_AXIS_MOVEMENT AT %I421.1 : Bool;
   Z_AXIS_MOVEMENT AT %I421.2 : Bool;
   R_AXIS_MOVEMENT AT %I421.3 : Bool;
   Z_ASIS_IN_ON_FOCUS AT %I421.4 : Bool;
   FOCUS_DISTANCE_SENSOR_IS_AVAILABLE AT %I421.5 : Bool;
   RESERVE_I_22_BYTE AT %IB422 : Byte;
   RESERVE_I_23_BYTE AT %IB423 : Byte;
   SET_OUTPUT AT %I424.0 : Bool;
   RESET_OUTPUT_IN AT %I424.1 : Bool;
   RRESERVE_I_25_BYTE AT %IB425 : Byte;
   I_O_PORT_LASER_OUTPUT_STATUS_0 AT %I426.0 : Bool;
   I_O_PORT_LASER_OUTPUT_STATUS_1 AT %I426.1 : Bool;
   I_O_PORT_LASER_OUTPUT_STATUS_2 AT %I426.2 : Bool;
   I_O_PORT_LASER_OUTPUT_STATUS_3 AT %I426.3 : Bool;
   I_O_PORT_LASER_OUTPUT_STATUS_4 AT %I426.4 : Bool;
   I_O_PORT_LASER_OUTPUT_STATUS_5 AT %I426.5 : Bool;
   I_O_PORT_LASER_OUTPUT_STATUS_6 AT %I426.6 : Bool;
   I_O_PORT_LASER_OUTPUT_STATUS_7 AT %I426.7 : Bool;
   I_O_PORT_LASER_OUTPUT_STATUS_8 AT %I427.0 : Bool;
   I_O_PORT_LASER_OUTPUT_STATUS_9 AT %I427.1 : Bool;
   I_O_PORT_LASER_OUTPUT_STATUS_10 AT %I427.2 : Bool;
   I_O_PORT_LASER_OUTPUT_STATUS_11 AT %I427.3 : Bool;
   I_O_PORT_LASER_OUTPUT_STATUS_12 AT %I427.4 : Bool;
   I_O_PORT_LASER_OUTPUT_STATUS_13 AT %I427.5 : Bool;
   I_O_PORT_LASER_OUTPUT_STATUS_14 AT %I427.6 : Bool;
   I_O_PORT_LASER_OUTPUT_STATUS_15 AT %I427.7 : Bool;
   I_O_PORT_LASER_INPUT_STATUS_0 AT %I428.0 : Bool;
   I_O_PORT_LASER_INPUT_STATUS_1 AT %I428.1 : Bool;
   I_O_PORT_LASER_INPUT_STATUS_2 AT %I428.2 : Bool;
   I_O_PORT_LASER_INPUT_STATUS_3 AT %I428.3 : Bool;
   I_O_PORT_LASER_INPUT_STATUS_4 AT %I428.4 : Bool;
   I_O_PORT_LASER_INPUT_STATUS_5 AT %I428.5 : Bool;
   I_O_PORT_LASER_INPUT_STATUS_6 AT %I428.6 : Bool;
   I_O_PORT_LASER_INPUT_STATUS_7 AT %I428.7 : Bool;
   I_O_PORT_LASER_INPUT_STATUS_8 AT %I429.0 : Bool;
   I_O_PORT_LASER_INPUT_STATUS_9 AT %I429.1 : Bool;
   I_O_PORT_LASER_INPUT_STATUS_10 AT %I429.2 : Bool;
   I_O_PORT_LASER_INPUT_STATUS_11 AT %I429.3 : Bool;
   I_O_PORT_LASER_INPUT_STATUS_12 AT %I429.4 : Bool;
   I_O_PORT_LASER_INPUT_STATUS_13 AT %I429.5 : Bool;
   I_O_PORT_LASER_INPUT_STATUS_14 AT %I429.6 : Bool;
   I_O_PORT_LASER_INPUT_STATUS_15 AT %I429.7 : Bool;
   RESERVE_I_30_BYTE AT %IB430 : Byte;
   RESERVE_I_31_BYTE AT %IB431 : Byte;
   RESERVE_I_32_BYTE AT %IB432 : Byte;
   RESERVE_I_33_BYTE AT %IB433 : Byte;
   GET_ID_MATCH_RESULT_IN AT %I434.1 : Bool;
   GET_ID_MARVIS_CONFIGURATION_IN AT %I434.2 : Bool;
   SET_ID_MARVIS_CONFIGURATION_IN AT %I434.3 : Bool;
   GET_ID_MARVIS_RESULT_IN AT %I434.4 : Bool;
   RESERVE_I_35_BYTE AT %IB435 : Byte;
   MARVIS_RESULT_OK AT %I436.0 : Bool;
   MARVIS_RESULT_FAIL AT %I436.1 : Bool;
   SYMBOL_READ_OK AT %I436.2 : Bool;
   SYMBOL_READ_FAIL AT %I436.3 : Bool;
   SYMBOL_GRADE_RESULT_OK AT %I436.4 : Bool;
   SYMBOL_GRADE_RESULT_FAIL AT %I436.5 : Bool;
   SYMBOL_MATCH_RESULT_OK AT %I436.6 : Bool;
   SYMBOL_MATCH_RESULT_FAIL AT %I436.7 : Bool;
   RESERVE_I_37_BYTE AT %IB437 : Byte;
   READER_STATUS_AVAILABLE AT %I438.1 : Bool;
   READER_STATUS_BZSY AT %I438.2 : Bool;
   READER_STATUS_WARNING AT %I438.3 : Bool;
   READER_STATUS_ERROR AT %I438.4 : Bool;
   RESERVE_I_39_BYTE AT %IB439 : Byte;
   RESERVE_I_40_BYTE AT %IB440 : Byte;
   RESERVE_I_41_BYTE AT %IB441 : Byte;
   RESERVE_I_42_BYTE AT %IB442 : Byte;
   RESERVE_I_43_BYTE AT %IB443 : Byte;
   RESERVE_I_44_BYTE AT %IB444 : Byte;
   RESERVE_I_45_BYTE AT %IB445 : Byte;
   RESERVE_I_46_BYTE AT %IB446 : Byte;
   RESERVE_I_47_BYTE AT %IB447 : Byte;
   RESERVE_I_48_BYTE AT %IB448 : Byte;
   RESERVE_I_49_BYTE AT %IB449 : Byte;
   RESERVE_I_50_BYTE AT %IB450 : Byte;
   RESERVE_I_51_BYTE AT %IB451 : Byte;
   RESERVE_I_52_BYTE AT %IB452 : Byte;
   RESERVE_I_53_BYTE AT %IB453 : Byte;
   RESPONSE_DATE_SIZE AT %IB454 : Byte;
   RESERVE_I_55_BYTE AT %IB455 : Byte;
   RESPONSE_DATA_FIELD_0 AT %IB456 : Byte;
   RESPONSE_DATA_FIELD_1 AT %IB457 : Byte;
   RESPONSE_DATA_FIELD_2 AT %IB458 : Byte;
   RESPONSE_DATA_FIELD_3 AT %IB459 : Byte;
   RESPONSE_DATA_FIELD_4 AT %IB460 : Byte;
   RESPONSE_DATA_FIELD_5 AT %IB461 : Byte;
   RESPONSE_DATA_FIELD_6 AT %IB462 : Byte;
   RESPONSE_DATA_FIELD_7 AT %IB463 : Byte;
   RESPONSE_DATA_FIELD_8 AT %IB464 : Byte;
   RESPONSE_DATA_FIELD_9 AT %IB465 : Byte;
   RESPONSE_DATA_FIELD_10 AT %IB466 : Byte;
   RESPONSE_DATA_FIELD_11 AT %IB467 : Byte;
   RESPONSE_DATA_FIELD_12 AT %IB468 : Byte;
   RESPONSE_DATA_FIELD_13 AT %IB469 : Byte;
   RESPONSE_DATA_FIELD_14 AT %IB470 : Byte;
   RESPONSE_DATA_FIELD_15 AT %IB471 : Byte;
   RESPONSE_DATA_FIELD_16 AT %IB472 : Byte;
   RESPONSE_DATA_FIELD_17 AT %IB473 : Byte;
   RESPONSE_DATA_FIELD_18 AT %IB474 : Byte;
   RESPONSE_DATA_FIELD_19 AT %IB475 : Byte;
   RESPONSE_DATA_FIELD_20 AT %IB476 : Byte;
   RESPONSE_DATA_FIELD_21 AT %IB477 : Byte;
   RESPONSE_DATA_FIELD_22 AT %IB478 : Byte;
   RESPONSE_DATA_FIELD_23 AT %IB479 : Byte;
   RESPONSE_DATA_FIELD_24 AT %IB480 : Byte;
   RESPONSE_DATA_FIELD_25 AT %IB481 : Byte;
   RESPONSE_DATA_FIELD_26 AT %IB482 : Byte;
   RESPONSE_DATA_FIELD_27 AT %IB483 : Byte;
   RESPONSE_DATA_FIELD_28 AT %IB484 : Byte;
   RESPONSE_DATA_FIELD_29 AT %IB485 : Byte;
   RESPONSE_DATA_FIELD_30 AT %IB486 : Byte;
   RESPONSE_DATA_FIELD_31 AT %IB487 : Byte;
   RESPONSE_DATA_FIELD_32 AT %IB488 : Byte;
   RESPONSE_DATA_FIELD_33 AT %IB489 : Byte;
   RESPONSE_DATA_FIELD_34 AT %IB490 : Byte;
   RESPONSE_DATA_FIELD_35 AT %IB491 : Byte;
   RESPONSE_DATA_FIELD_36 AT %IB492 : Byte;
   RESPONSE_DATA_FIELD_37 AT %IB493 : Byte;
   RESPONSE_DATA_FIELD_38 AT %IB494 : Byte;
   RESPONSE_DATA_FIELD_39 AT %IB495 : Byte;
   RESPONSE_DATA_FIELD_40 AT %IB496 : Byte;
   RESPONSE_DATA_FIELD_41 AT %IB497 : Byte;
   RESPONSE_DATA_FIELD_42 AT %IB498 : Byte;
   RESPONSE_DATA_FIELD_43 AT %IB499 : Byte;
   RESPONSE_DATA_FIELD_44 AT %IB500 : Byte;
   RESPONSE_DATA_FIELD_45 AT %IB501 : Byte;
   RESPONSE_DATA_FIELD_46 AT %IB502 : Byte;
   RESPONSE_DATA_FIELD_47 AT %IB503 : Byte;
   RESPONSE_DATA_FIELD_48 AT %IB504 : Byte;
   RESPONSE_DATA_FIELD_49 AT %IB505 : Byte;
   RESPONSE_DATA_FIELD_50 AT %IB506 : Byte;
   RESPONSE_DATA_FIELD_51 AT %IB507 : Byte;
   RESPONSE_DATA_FIELD_52 AT %IB508 : Byte;
   RESPONSE_DATA_FIELD_53 AT %IB509 : Byte;
   RESPONSE_DATA_FIELD_54 AT %IB510 : Byte;
   RESPONSE_DATA_FIELD_55 AT %IB511 : Byte;
   RESPONSE_DATA_FIELD_56 AT %IB512 : Byte;
   RESPONSE_DATA_FIELD_57 AT %IB513 : Byte;
   RESPONSE_DATA_FIELD_58 AT %IB514 : Byte;
   RESPONSE_DATA_FIELD_59 AT %IB515 : Byte;
   RESPONSE_DATA_FIELD_60 AT %IB516 : Byte;
   RESPONSE_DATA_FIELD_61 AT %IB517 : Byte;
   RESPONSE_DATA_FIELD_62 AT %IB518 : Byte;
   RESPONSE_DATA_FIELD_63 AT %IB519 : Byte;
   RESPONSE_DATA_FIELD_64 AT %IB520 : Byte;
   RESPONSE_DATA_FIELD_65 AT %IB521 : Byte;
   RESPONSE_DATA_FIELD_66 AT %IB522 : Byte;
   RESPONSE_DATA_FIELD_67 AT %IB523 : Byte;
   RESPONSE_DATA_FIELD_68 AT %IB524 : Byte;
   RESPONSE_DATA_FIELD_69 AT %IB525 : Byte;
   RESPONSE_DATA_FIELD_70 AT %IB526 : Byte;
   RESPONSE_DATA_FIELD_71 AT %IB527 : Byte;
END_VAR

VAR_GLOBAL   // PLC tag table "LASER_OUT_datalogic"
   START_MARKING AT %Q1500.0 : Bool;
   STOP_SYSTEM AT %Q1500.1 : Bool;
   GET_PNIO_PROTOCOL_VERSION AT %Q1501.0 : Bool;
   PROTOCOL_ERROR_CLEAR AT %Q1501.7 : Bool;
   OPEN_DOKUMENT_FROM_DEVICE AT %Q1502.0 : Bool;
   SAVE_DOKUMENT AT %Q1502.1 : Bool;
   GET_DATA_FIELD_VALUE AT %Q1502.2 : Bool;
   SET_DATA_FIELD_VALUE AT %Q1502.3 : Bool;
   GET_GLOBAL_COUNTER_VALUE AT %Q1502.4 : Bool;
   SET_GLOBAL_COUNTER_VALUE AT %Q1502.5 : Bool;
   GET_GLOBAL_STRING_VALUE AT %Q1502.6 : Bool;
   SET_GLOBAL_STRING_VALUE AT %Q1502.7 : Bool;
   ENABLE_DATA_FIELD AT %Q1503.0 : Bool;
   DISABLE_DATA_FIELD AT %Q1503.1 : Bool;
   MOVE_AND_ROTATE_DOCUMENT AT %Q1504.0 : Bool;
   MOVE_DATA_FIELD AT %Q1504.1 : Bool;
   RESERVE_Q_5_BYTE AT %QB1505 : Byte;
   RESERVE_Q_6_BYTE AT %QB1506 : Byte;
   RESERVE_Q_7_BYTE AT %QB1507 : Byte;
   MOVE_AXIS AT %Q1508.0 : Bool;
   RESET_AXIS AT %Q1508.1 : Bool;
   STOP_AXIS AT %Q1508.2 : Bool;
   START_AUTOFOCUS AT %Q1508.3 : Bool;
   STOP_AUTOFOCUS AT %Q1508.4 : Bool;
   SET_FOCUS_DISTANCE_SENSOR_REFERENCE AT %Q1508.5 : Bool;
   RESERVE_Q_9_BYTE AT %QB1509 : Byte;
   X_AXIS AT %Q1510.0 : Bool;
   Y_AXIS AT %Q1510.1 : Bool;
   Z_AXIS AT %Q1510.2 : Bool;
   R_AXIS AT %Q1510.3 : Bool;
   RESERVE_Q_11_BYTE AT %QB411 : Byte;
   RESERVE_Q_12_BYTE AT %QB412 : Byte;
   RESERVE_Q_13_BYTE AT %QB413 : Byte;
   RESERVE_Q_14_BYTE AT %QB414 : Byte;
   RESERVE_Q_15_BYTE AT %QB415 : Byte;
   RESERVE_Q_16_BYTE AT %QB416 : Byte;
   RESERVE_Q_17_BYTE AT %QB417 : Byte;
   RESERVE_Q_18_BYTE AT %QB418 : Byte;
   RESERVE_Q_19_BYTE AT %QB419 : Byte;
   RESERVE_Q_20_BYTE AT %QB420 : Byte;
   RESERVE_Q_21_BYTE AT %QB421 : Byte;
   SET_AUTPUT AT %Q1522.0 : Bool;
   RESET_OUTPUT AT %Q1522.1 : Bool;
   RESERVE_Q_23_BYTE AT %QB1523 : Byte;   // --------------------
   I_O_PORT_LASER_OUTPUT_0 AT %Q1524.0 : Bool;
   I_O_PORT_LASER_OUTPUT_1 AT %Q1524.1 : Bool;
   I_O_PORT_LASER_OUTPUT_2 AT %Q1524.2 : Bool;
   I_O_PORT_LASER_OUTPUT_3 AT %Q1524.3 : Bool;
   I_O_PORT_LASER_OUTPUT_4 AT %Q1524.4 : Bool;
   I_O_PORT_LASER_OUTPUT_5 AT %Q1524.5 : Bool;
   I_O_PORT_LASER_OUTPUT_6 AT %Q1524.6 : Bool;
   I_O_PORT_LASER_OUTPUT_7 AT %Q1524.7 : Bool;
   I_O_PORT_LASER_OUTPUT_8 AT %Q1525.0 : Bool;
   I_O_PORT_LASER_OUTPUT_9 AT %Q1525.1 : Bool;
   I_O_PORT_LASER_OUTPUT_10 AT %Q1525.2 : Bool;
   I_O_PORT_LASER_OUTPUT_11 AT %Q1525.3 : Bool;
   I_O_PORT_LASER_OUTPUT_12 AT %Q1525.4 : Bool;
   I_O_PORT_LASER_OUTPUT_13 AT %Q1525.5 : Bool;
   I_O_PORT_LASER_OUTPUT_14 AT %Q1525.6 : Bool;
   I_O_PORT_LASER_OUTPUT_15 AT %Q1525.7 : Bool;
   RESERVE_Q_26_BYTE AT %QB1526 : Byte;   // --------------------
   RESERVE_Q_27_BYTE AT %QB1527 : Byte;   // --------------------
   RESERVE_Q_28_BYTE AT %QB1528 : Byte;   // --------------------
   RESERVE_Q_29_BYTE AT %QB1529 : Byte;   // --------------------
   RESERVE_Q_30_BYTE AT %QB1530 : Byte;   // --------------------
   RESERVE_Q_31_BYTE AT %QB1531 : Byte;   // --------------------
   GET_ID_MATCH_RESULT AT %Q1532.1 : Bool;
   GET_ID_MARVIS_CONFIGURATION AT %Q1532.2 : Bool;
   SET_ID_MARVIS_CONFIGURATION AT %Q1532.3 : Bool;
   GET_ID_MARVIS_RESULT AT %Q1532.4 : Bool;
   RESERVE_Q_33_BYTE AT %QB1533 : Byte;
   RESERVE_Q_34_BYTE AT %QB1534 : Byte;
   RESERVE_Q_35_BYTE AT %QB1535 : Byte;
   RESERVE_Q_36_BYTE AT %QB1536 : Byte;
   RESERVE_Q_37_BYTE AT %QB1537 : Byte;
   RESERVE_Q_38_BYTE AT %QB1538 : Byte;
   RESERVE_Q_39_BYTE AT %QB1539 : Byte;
   RESERVE_Q_40_BYTE AT %QB1540 : Byte;
   RESERVE_Q_41_BYTE AT %QB1541 : Byte;
   RESERVE_Q_42_BYTE AT %QB1542 : Byte;
   RESERVE_Q_43_BYTE AT %QB1543 : Byte;
   RESERVE_Q_44_BYTE AT %QB1544 : Byte;
   RESERVE_Q_45_BYTE AT %QB1545 : Byte;
   RESERVE_Q_46_BYTE AT %QB1546 : Byte;
   RESERVE_Q_47_BYTE AT %QB1547 : Byte;
   RESERVE_Q_48_BYTE AT %QB1548 : Byte;
   RESERVE_Q_49_BYTE AT %QB1549 : Byte;
   RESERVE_Q_50_BYTE AT %QB1550 : Byte;
   RESERVE_Q_51_BYTE AT %QB1551 : Byte;
   RESERVE_Q_52_BYTE AT %QB1552 : Byte;
   RESERVE_Q_53_BYTE AT %QB1553 : Byte;
   REQUEST_DATA_SIZE AT %QB1554 : Byte;
   RESERVE_Q_55_BYTE AT %QB1555 : Byte;
   REQUEST_DATA_FIELC_BYTE_0 AT %QB1556 : Byte;
   REQUEST_DATA_FIELC_BYTE_1 AT %QB1557 : Byte;
   REQUEST_DATA_FIELC_BYTE_2 AT %QB1558 : Byte;
   REQUEST_DATA_FIELC_BYTE_3 AT %QB1559 : Byte;
   REQUEST_DATA_FIELC_BYTE_4 AT %QB1560 : Byte;
   REQUEST_DATA_FIELC_BYTE_5 AT %QB1561 : Byte;
   REQUEST_DATA_FIELC_BYTE_6 AT %QB1562 : Byte;
   REQUEST_DATA_FIELC_BYTE_7 AT %QB1563 : Byte;
   REQUEST_DATA_FIELC_BYTE_8 AT %QB1564 : Byte;
   REQUEST_DATA_FIELC_BYTE_9 AT %QB1565 : Byte;
   REQUEST_DATA_FIELC_BYTE_10 AT %QB1566 : Byte;
   REQUEST_DATA_FIELC_BYTE_11 AT %QB1567 : Byte;
   REQUEST_DATA_FIELC_BYTE_12 AT %QB1568 : Byte;
   REQUEST_DATA_FIELC_BYTE_13 AT %QB1569 : Byte;
   REQUEST_DATA_FIELC_BYTE_14 AT %QB1570 : Byte;
   REQUEST_DATA_FIELC_BYTE_15 AT %QB1571 : Byte;
   REQUEST_DATA_FIELC_BYTE_16 AT %QB1572 : Byte;
   REQUEST_DATA_FIELC_BYTE_17 AT %QB1573 : Byte;
   REQUEST_DATA_FIELC_BYTE_18 AT %QB1574 : Byte;
   REQUEST_DATA_FIELC_BYTE_19 AT %QB1575 : Byte;
   REQUEST_DATA_FIELC_BYTE_20 AT %QB1576 : Byte;
   REQUEST_DATA_FIELC_BYTE_21 AT %QB1577 : Byte;
   REQUEST_DATA_FIELC_BYTE_22 AT %QB1578 : Byte;
   REQUEST_DATA_FIELC_BYTE_23 AT %QB1579 : Byte;
   REQUEST_DATA_FIELC_BYTE_24 AT %QB1580 : Byte;
   REQUEST_DATA_FIELC_BYTE_25 AT %QB1581 : Byte;
   REQUEST_DATA_FIELC_BYTE_26 AT %QB1582 : Byte;
   REQUEST_DATA_FIELC_BYTE_27 AT %QB1583 : Byte;
   REQUEST_DATA_FIELC_BYTE_28 AT %QB1584 : Byte;
   REQUEST_DATA_FIELC_BYTE_29 AT %QB1585 : Byte;
   REQUEST_DATA_FIELC_BYTE_30 AT %QB1586 : Byte;
   REQUEST_DATA_FIELC_BYTE_31 AT %QB1587 : Byte;
   REQUEST_DATA_FIELC_BYTE_32 AT %QB1588 : Byte;
   REQUEST_DATA_FIELC_BYTE_33 AT %QB1589 : Byte;
   REQUEST_DATA_FIELC_BYTE_34 AT %QB1590 : Byte;
   REQUEST_DATA_FIELC_BYTE_35 AT %QB1591 : Byte;
   REQUEST_DATA_FIELC_BYTE_36 AT %QB1592 : Byte;
   REQUEST_DATA_FIELC_BYTE_37 AT %QB1593 : Byte;
   REQUEST_DATA_FIELC_BYTE_38 AT %QB1594 : Byte;
   REQUEST_DATA_FIELC_BYTE_39 AT %QB1595 : Byte;
   REQUEST_DATA_FIELC_BYTE_40 AT %QB1596 : Byte;
   REQUEST_DATA_FIELC_BYTE_41 AT %QB1597 : Byte;
   REQUEST_DATA_FIELC_BYTE_42 AT %QB1598 : Byte;
   REQUEST_DATA_FIELC_BYTE_43 AT %QB1599 : Byte;
   REQUEST_DATA_FIELC_BYTE_44 AT %QB1600 : Byte;
   REQUEST_DATA_FIELC_BYTE_45 AT %QB1601 : Byte;
   REQUEST_DATA_FIELC_BYTE_46 AT %QB1602 : Byte;
   REQUEST_DATA_FIELC_BYTE_47 AT %QB1603 : Byte;
   REQUEST_DATA_FIELC_BYTE_48 AT %QB1604 : Byte;
   REQUEST_DATA_FIELC_BYTE_49 AT %QB1605 : Byte;
   REQUEST_DATA_FIELC_BYTE_50 AT %QB1606 : Byte;
   REQUEST_DATA_FIELC_BYTE_51 AT %QB1607 : Byte;
   REQUEST_DATA_FIELC_BYTE_52 AT %QB1608 : Byte;
   REQUEST_DATA_FIELC_BYTE_53 AT %QB1609 : Byte;
   REQUEST_DATA_FIELC_BYTE_54 AT %QB1610 : Byte;
   REQUEST_DATA_FIELC_BYTE_55 AT %QB1611 : Byte;
   REQUEST_DATA_FIELC_BYTE_56 AT %QB1612 : Byte;
   REQUEST_DATA_FIELC_BYTE_57 AT %QB1613 : Byte;
   REQUEST_DATA_FIELC_BYTE_58 AT %QB1614 : Byte;
   REQUEST_DATA_FIELC_BYTE_59 AT %QB1615 : Byte;
   REQUEST_DATA_FIELC_BYTE_60 AT %QB1616 : Byte;
   REQUEST_DATA_FIELC_BYTE_61 AT %QB1617 : Byte;
   REQUEST_DATA_FIELC_BYTE_62 AT %QB1618 : Byte;
   REQUEST_DATA_FIELC_BYTE_63 AT %QB1619 : Byte;
   REQUEST_DATA_FIELC_BYTE_64 AT %QB1620 : Byte;
   REQUEST_DATA_FIELC_BYTE_65 AT %QB1621 : Byte;
   REQUEST_DATA_FIELC_BYTE_66 AT %QB1622 : Byte;
   REQUEST_DATA_FIELC_BYTE_67 AT %QB1623 : Byte;
   REQUEST_DATA_FIELC_BYTE_68 AT %QB1624 : Byte;
   REQUEST_DATA_FIELC_BYTE_69 AT %QB1625 : Byte;
   REQUEST_DATA_FIELC_BYTE_70 AT %QB1626 : Byte;
   REQUEST_DATA_FIELC_BYTE_71 AT %QB1627 : Byte;
END_VAR

VAR_GLOBAL   // PLC tag table "Laser_in_macsa"
   "-XT500_d_counter" AT %ID1583 : DWord;   // counter indicating the number of o.k. prints since entering into the printing mode
   "-XT500_s_counter" AT %ID1587 : DWord;   // counter indicating the number of prints since entering into the printing mode.
   "-XT500_messageport" AT %ID1591 : DWord;   // indicates the bit combination of the external message selection (when external message mode is activated)
   "-XT500_status_byte_0" AT %IB1595 : Byte;
   "-XT500_status_byte_1" AT %IB1596 : Byte;   // 0x00: default value. -- 0x01: request; the system is requesting information to
   "-XT500_status_byte_2" AT %IB1597 : Byte;   // option byte; (internal use), indicates the type of
   "-XT500_status_byte_3" AT %IB1598 : Byte;   // 0x00: default , system is in standard mode. 0x01: system is in external message selection mode 0x04: system is in a batch-job mode.
   "-XT500_t_counter" AT %ID1599 : DWord;   // 32-bit counter indicating the total number of prints of the laser system
   "-XT500_copies" AT %ID1603 : DWord;   // the actual number of print copies.
   "-XT500_alarm_information" AT %IW1609 : Word;   // 0X0000: no alarms -- 0x0C0E: wrong messageport (no file found for the external message selection) -- 0x0848: alarms active; some alarms are active (interlock, shutter,....) -- 0xFFFF: initialization of the firmware has failed due to some hardware failure.
   "-XT500_prinntime" AT %ID1611 : DWord;   // print time
   "-XT500_alarm-mask" AT %ID1616 : DWord;   // popis panel text end grafik list
   "-XT500_signalstate" AT %ID1619 : DWord;
   "-XT500_name_byte_0" AT %IB1623 : Byte;   // actual filename + extension of the message.
   "-XT500_name_byte_1" AT %IB1624 : Byte;   // actual filename + extension of the message.
   "-XT500_name_byte_2" AT %IB1625 : Byte;   // actual filename + extension of the message.
   "-XT500_name_byte_3" AT %IB1626 : Byte;   // actual filename + extension of the message.
   "-XT500_name_byte_4" AT %IB1627 : Byte;   // actual filename + extension of the message.
   "-XT500_name_byte_5" AT %IB1628 : Byte;   // actual filename + extension of the message.
   "-XT500_name_byte_6" AT %IB1629 : Byte;   // actual filename + extension of the message.
   "-XT500_name_byte_7" AT %IB1630 : Byte;   // actual filename + extension of the message.
   "-XT500_name_byte_8" AT %IB1631 : Byte;   // actual filename + extension of the message.
   "-XT500_name_byte_9" AT %IB1632 : Byte;   // actual filename + extension of the message.
   "-XT500_name_byte_10" AT %IB1633 : Byte;   // actual filename + extension of the message.
   "-XT500_name_byte_11" AT %IB1634 : Byte;   // actual filename + extension of the message.
   "-XT500_name_byte_12" AT %IB1635 : Byte;   // actual filename + extension of the message.
   "-XT500_name_byte_13" AT %IB1636 : Byte;   // actual filename + extension of the message.
   "-XT500_name_byte_14" AT %IB1637 : Byte;   // actual filename + extension of the message.
   "-XT500_name_byte_15" AT %IB1638 : Byte;   // actual filename + extension of the message.
   "-XT500_eventhandler_byte_0" AT %IB1639 : Byte;   // actual filename + extension of the eventhandler-file.
   "-XT500_eventhandler_byte_1" AT %IB1640 : Byte;   // actual filename + extension of the eventhandler-file.
   "-XT500_eventhandler_byte_2" AT %IB1641 : Byte;   // actual filename + extension of the eventhandler-file.
   "-XT500_eventhandler_byte_3" AT %IB1642 : Byte;   // actual filename + extension of the eventhandler-file.
   "-XT500_eventhandler_byte_4" AT %IB1643 : Byte;   // actual filename + extension of the eventhandler-file.
   "-XT500_eventhandler_byte_5" AT %IB1644 : Byte;   // actual filename + extension of the eventhandler-file.
   "-XT500_eventhandler_byte_6" AT %IB1645 : Byte;   // actual filename + extension of the eventhandler-file.
   "-XT500_eventhandler_byte_7" AT %IB1646 : Byte;   // actual filename + extension of the eventhandler-file.
   "-XT500_eventhandler_byte_8" AT %IB1647 : Byte;   // actual filename + extension of the eventhandler-file.
   "-XT500_eventhandler_byte_9" AT %IB1648 : Byte;   // actual filename + extension of the eventhandler-file.
   "-XT500_eventhandler_byte_10" AT %IB1649 : Byte;   // actual filename + extension of the eventhandler-file.
   "-XT500_eventhandler_byte_11" AT %IB1650 : Byte;   // actual filename + extension of the eventhandler-file.
   "-XT500_eventhandler_byte_12" AT %IB1651 : Byte;   // actual filename + extension of the eventhandler-file.
   "-XT500_eventhandler_byte_13" AT %IB1652 : Byte;   // actual filename + extension of the eventhandler-file.
   "-XT500_eventhandler_byte_14" AT %IB1653 : Byte;   // actual filename + extension of the eventhandler-file.
   "-XT500_eventhandler_byte_15" AT %IB1654 : Byte;   // actual filename + extension of the eventhandler-file.
   "-XT500_extended_alarm-mask" AT %ID1655 : DWord;   // See Status command. When the alarm-mask has the ‘extended alarmmask’ rozepsano text list
   "-XT500_not_used_0" AT %IB1659 : Byte;
   "-XT500_not_used_1" AT %IB1660 : Byte;
   "-XT500_scanfield_0" AT %IB1661 : Byte;
   "-XT500_scanfield_1" AT %IB1662 : Byte;
   "-XT500_data_recived_byte" AT %IB1663 : Byte;   // status
   "-XT500_data_recived_byte_0" AT %I1663.0 : Bool;   // data ready
   "-XT500_data_recived_byte_1" AT %I1663.1 : Bool;   // clear command error trigger
   "-XT500_data_recived_byte_2" AT %I1663.2 : Bool;
   "-XT500_data_recived_byte_3" AT %I1663.3 : Bool;
   "-XT500_data_recived_byte_4" AT %I1663.4 : Bool;
   "-XT500_data_recived_byte_5" AT %I1663.5 : Bool;
   "-XT500_data_recived_byte_6" AT %I1663.6 : Bool;
   "-XT500_data_recived_byte_7" AT %I1663.7 : Bool;
   "-XT500_command_error_info" AT %IW1664 : Word;   // command error info (0xFF == command
   "-XT500_status_byte_0_bool_0" AT %I1595.0 : Bool;   // when set, system is in printing mode (waiting for photocell/PLC)
   "-XT500_status_byte_0_bool_1" AT %I1595.1 : Bool;   // when set, system is actually printing a message
   "-XT500_status_byte_0_bool_2" AT %I1595.2 : Bool;   // when set, system is waiting for a 'alarm reset' signal (DSP cards only).
   "-XT500_status_byte_0_bool_3" AT %I1595.3 : Bool;   // when set, system is waiting for an input signal (DSP cards only)
   "-XT500_status_byte_0_bool_4" AT %I1595.4 : Bool;   // when set, system is waiting for an external motorized axis to reach a new position.
   "-XT500_status_byte_0_bool_5" AT %I1595.5 : Bool;   // when set, system is in ‘printsession’ mode.
   "-XT500_status_byte_0_bool_6" AT %I1595.6 : Bool;   // reserved
   "-XT500_status_byte_0_bool_7" AT %I1595.7 : Bool;   // reserved
   "-XT500_status_byte_1_bool_0" AT %I1596.0 : Bool;
   "-XT500_status_byte_1_bool_1" AT %I1596.1 : Bool;
   "-XT500_status_byte_1_bool_2" AT %I1596.2 : Bool;
   "-XT500_status_byte_1_bool_3" AT %I1596.3 : Bool;
   "-XT500_status_byte_1_bool_4" AT %I1596.4 : Bool;
   "-XT500_status_byte_1_bool_5" AT %I1596.5 : Bool;
   "-XT500_status_byte_1_bool_6" AT %I1596.6 : Bool;
   "-XT500_status_byte_1_bool_7" AT %I1596.7 : Bool;
   "-XT500_scanfield_1_bit_8" AT %I1662.0 : Bool;
   "-XT500_scanfield_1_bit_9" AT %I1662.1 : Bool;
   "-XT500_scanfield_1_bit_10" AT %I1662.2 : Bool;   // 0: static
   "-XT500_scanfield_1_bit_11" AT %I1662.3 : Bool;   // 1: dynamic
   "-XT500_scanfield_1_bit_12" AT %I1662.4 : Bool;   // 2: dynamic-distance
   "-XT500_scanfield_1_bit_13" AT %I1662.5 : Bool;   // 3: static-dynamic
   "-XT500_scanfield_1_bit_14" AT %I1662.6 : Bool;   // 4: stepper mode
   "-XT500_scanfield_1_bit_15" AT %I1662.7 : Bool;   // 5: XY stepper mode
   "-XT500_alarm-mask_interlock" AT %I1618.0 : Bool;   // interlock součást alarm-mask
   "-XT500_alarm-mask_shutter" AT %I1618.3 : Bool;   // shutter součást alarm-mask oim
   "-XT500_alarm-mask_laser_not_ready" AT %I1618.4 : Bool;   // laser nor ready součást alarm mask
   "-XT500_alarm-mask_laser_not_armed" AT %I1619.3 : Bool;   // laser nor armed součást alarm mask
   "-XT500_alarm_mas_warm_up_in_progres" AT %I1619.5 : Bool;   // warm_up_in_progres součást alarm mask
   "-XT500_alarm-mask_shutter_oim" AT %I1618.1 : Bool;
   "-XT500_copies_1" AT %IW1605 : Word;
   "-XT500_copies_2" AT %IW1607 : Word;
   "-XT500_Tag_1" AT %I1618.2 : Bool;
   "-XT500_alarm_information(1)" AT %IW1610 : Word;   // 0X0000: no alarms -- 0x0C0E: wrong messageport (no file found for the external message selection) -- 0x0848: alarms active; some alarms are active (interlock, shutter,....) -- 0xFFFF: initialization of the firmware has failed due to some hardware failure.
   "-XT500_alarm_information(2)" AT %IW1608 : Word;   // 0X0000: no alarms -- 0x0C0E: wrong messageport (no file found for the external message selection) -- 0x0848: alarms active; some alarms are active (interlock, shutter,....) -- 0xFFFF: initialization of the firmware has failed due to some hardware failure.
   "-XT500_alarm_information(3)" AT %IW1611 : Word;   // 0X0000: no alarms -- 0x0C0E: wrong messageport (no file found for the external message selection) -- 0x0848: alarms active; some alarms are active (interlock, shutter,....) -- 0xFFFF: initialization of the firmware has failed due to some hardware failure.
   "-XT500_alarm_information_bool_1" AT %I1610.0 : Bool;
   "-XT500_alarm_information_bool_2" AT %I1610.1 : Bool;
   "-XT500_alarm_information_bool_3" AT %I1610.2 : Bool;
   "-XT500_alarm_information_bool_4" AT %I1610.3 : Bool;   // neni_nahrato_1
   "-XT500_alarm_information_bool_5" AT %I1610.4 : Bool;
   "-XT500_alarm_information_bool_6" AT %I1610.5 : Bool;
   "-XT500_alarm_information_bool_7" AT %I1610.6 : Bool;   // neni_najrato_2
   "-XT500_alarm_information_bool_8" AT %I1610.7 : Bool;
END_VAR

VAR_GLOBAL   // PLC tag table "laser_out_macsa"
   "-XT500_output_mode" AT %QD295 : DWord;   // Pole - výber pole podle čísla max 255
   "-XT500_output_byte_1" AT %QB295 : Byte;
   "-XT500_output_byte_2" AT %QB296 : Byte;
   "-XT500_output_byte_3" AT %QB297 : Byte;
   "-XT500_output_byte_4" AT %QB298 : Byte;
   "-XT500_output_copies" AT %QD299 : DWord;
   "-XT500_output_byte_5" AT %QB299 : Byte;   // zapisovaná data
   "-XT500_output_byte_6" AT %QB300 : Byte;   // zapisovaná data
   "-XT500_output_byte_7" AT %QB301 : Byte;   // zapisovaná data
   "-XT500_output_byte_8" AT %QB302 : Byte;   // zapisovaná data
   "-XT500_output_byte_9" AT %QB303 : Byte;   // zapisovaná data
   "-XT500_output_batch" AT %QD303 : DWord;
   "-XT500_output_byte_10" AT %QB304 : Byte;   // zapisovaná data
   "-XT500_output_byte_11" AT %QB305 : Byte;   // zapisovaná data
   "-XT500_output_byte_12" AT %QB306 : Byte;   // zapisovaná data
   "-XT500_output_filename_1" AT %QB307 : Byte;   // zápid textu v asci pro volbu programu + další data
   "-XT500_output_filename_2" AT %QB308 : Byte;   // zápid textu v asci pro volbu programu + další data
   "-XT500_output_filename_3" AT %QB309 : Byte;   // zápid textu v asci pro volbu programu + další data
   "-XT500_output_filename_4" AT %QB310 : Byte;   // zápid textu v asci pro volbu programu + další data
   "-XT500_output_filename_5" AT %QB311 : Byte;   // zápid textu v asci pro volbu programu + další data
   "-XT500_output_filename_6" AT %QB312 : Byte;   // zápid textu v asci pro volbu programu + další data
   "-XT500_output_filename_7" AT %QB313 : Byte;   // zápid textu v asci pro volbu programu + další data
   "-XT500_output_filename_8" AT %QB314 : Byte;   // zápid textu v asci pro volbu programu + další data
   "-XT500_output_filename_9" AT %QB315 : Byte;   // zápid textu v asci pro volbu programu + další data
   "-XT500_output_filename_10" AT %QB316 : Byte;   // zápid textu v asci pro volbu programu + další data
   "-XT500_output_filename_11" AT %QB317 : Byte;   // zápid textu v asci pro volbu programu + další data
   "-XT500_output_filename_12" AT %QB318 : Byte;   // zápid textu v asci pro volbu programu + další data
   "-XT500_output_filename_13" AT %QB319 : Byte;   // zápid textu v asci pro volbu programu + další data
   "-XT500_output_filename_14" AT %QB320 : Byte;   // zápid textu v asci pro volbu programu + další data
   "-XT500_output_filename_15" AT %QB321 : Byte;   // zápid textu v asci pro volbu programu + další data
   "-XT500_output_filename_16" AT %QB322 : Byte;   // zápid textu v asci pro volbu programu + další data
   "-XT500_output_filename_17" AT %QB323 : Byte;   // zápid textu v asci pro volbu programu + další data
   "-XT500_command_number" AT %QB293 : Byte;   // výběr daného komandu v podobě čísla podle návodu zadavano v decu pozor na převod mezi word a int ----------- 6 zapis dat 16 vypal 1 otevření zprávy
   "-XT500_command_triger" AT %QB294 : Byte;   // 1= proveď příkaz
   "-XT500_output_filename_18" AT %QB324 : Byte;   // zápid textu v asci pro volbu programu + další data
   "-XT500_output_filename_19" AT %QB325 : Byte;   // zápid textu v asci pro volbu programu + další data
   "-XT500_output_filename_20" AT %QB326 : Byte;   // zápid textu v asci pro volbu programu + další data
   "-XT500_output_filename_21" AT %QB327 : Byte;   // zápid textu v asci pro volbu programu + další data
   "-XT500_output_filename_22" AT %QB328 : Byte;   // zápid textu v asci pro volbu programu + další data
   "-XT500_output_filename_23" AT %QB329 : Byte;   // zápid textu v asci pro volbu programu + další data
   "-XT500_output_filename_24" AT %QB330 : Byte;   // zápid textu v asci pro volbu programu + další data
   "-XT500_output_filename_25" AT %QB331 : Byte;   // zápid textu v asci pro volbu programu + další data
   "-XT500_output_filename_26" AT %QB332 : Byte;   // zápid textu v asci pro volbu programu + další data
   "-XT500_output_filename_27" AT %QB333 : Byte;   // zápid textu v asci pro volbu programu + další data
   "-XT500_output_filename_28" AT %QB334 : Byte;   // zápid textu v asci pro volbu programu + další data
   "-XT500_output_filename_29" AT %QB335 : Byte;   // zápid textu v asci pro volbu programu + další data
   "-XT500_output_filename_30" AT %QB336 : Byte;   // zápid textu v asci pro volbu programu + další data
   "-XT500_output_filename_31" AT %QB337 : Byte;   // zápid textu v asci pro volbu programu + další data
   "-XT500_output_filename_32" AT %QB338 : Byte;   // zápid textu v asci pro volbu programu + další data
   "-XT500_output_filename_33" AT %QB339 : Byte;   // zápid textu v asci pro volbu programu + další data
   "-XT500_output_filename_34" AT %QB340 : Byte;   // zápid textu v asci pro volbu programu + další data
   "-XT500_output_filename_35" AT %QB341 : Byte;   // zápid textu v asci pro volbu programu + další data
   "-XT500_output_filename_36" AT %QB342 : Byte;   // zápid textu v asci pro volbu programu + další data
   "-XT500_output_filename_37" AT %QB343 : Byte;   // zápid textu v asci pro volbu programu + další data
   "-XT500_output_filename_38" AT %QB344 : Byte;   // zápid textu v asci pro volbu programu + další data
   "-XT500_output_filename_39" AT %QB345 : Byte;   // zápid textu v asci pro volbu programu + další data
   "-XT500_output_filename_40" AT %QB346 : Byte;   // zápid textu v asci pro volbu programu + další data
   "-XT500_output_filename_41" AT %QB347 : Byte;   // zápid textu v asci pro volbu programu + další data
   "-XT500_output_filename_42" AT %QB348 : Byte;   // zápid textu v asci pro volbu programu + další data
   "-XT500_output_filename_43" AT %QB349 : Byte;   // zápid textu v asci pro volbu programu + další data
   "-XT500_output_filename_44" AT %QB350 : Byte;   // zápid textu v asci pro volbu programu + další data
   "-XT500_output_filename_45" AT %QB351 : Byte;   // zápid textu v asci pro volbu programu + další data
   "-XT500_output_filename_46" AT %QB352 : Byte;   // zápid textu v asci pro volbu programu + další data
   "-XT500_output_filename_47" AT %QB353 : Byte;   // zápid textu v asci pro volbu programu + další data
   "-XT500_output_filename_48" AT %QB354 : Byte;   // zápid textu v asci pro volbu programu + další data
   "-XT500_output_filename_49" AT %QB355 : Byte;   // zápid textu v asci pro volbu programu + další data
   "-XT500_output_filename_50" AT %QB356 : Byte;   // zápid textu v asci pro volbu programu + další data
   "-XT500_output_filename_51" AT %QB357 : Byte;   // zápid textu v asci pro volbu programu + další data
   "-XT500_output_filename_52" AT %QB358 : Byte;   // zápid textu v asci pro volbu programu + další data
   "-XT500_output_filename_53" AT %QB359 : Byte;   // zápid textu v asci pro volbu programu + další data
   "-XT500_output_filename_54" AT %QB360 : Byte;   // zápid textu v asci pro volbu programu + další data
   "-XT500_output_filename_55" AT %QB361 : Byte;   // zápid textu v asci pro volbu programu + další data
   "-XT500_output_filename_56" AT %QB362 : Byte;   // zápid textu v asci pro volbu programu + další data
   "-XT500_output_filename_57" AT %QB363 : Byte;   // zápid textu v asci pro volbu programu + další data
   "-XT500_output_filename_58" AT %QB364 : Byte;   // zápid textu v asci pro volbu programu + další data
   "-XT500_output_filename_59" AT %QB365 : Byte;   // zápid textu v asci pro volbu programu + další data
   "-XT500_output_filename_60" AT %QB366 : Byte;   // zápid textu v asci pro volbu programu + další data
   "-XT500_output_filename_61" AT %QB367 : Byte;   // zápid textu v asci pro volbu programu + další data
   "-XT500_output_filename_62" AT %QB368 : Byte;   // zápid textu v asci pro volbu programu + další data
   "-XT500_output_filename_63" AT %QB369 : Byte;   // zápid textu v asci pro volbu programu + další data
   "-XT500_output_filename_64" AT %QB370 : Byte;   // zápid textu v asci pro volbu programu + další data
   "-XT500_output_filename_65" AT %QB371 : Byte;   // zápid textu v asci pro volbu programu + další data
   "-XT500_output_filename_66" AT %QB372 : Byte;   // zápid textu v asci pro volbu programu + další data
   "-XT500_output_filename_67" AT %QB373 : Byte;   // zápid textu v asci pro volbu programu + další data
   "-XT500_output_filename_68" AT %QB374 : Byte;   // zápid textu v asci pro volbu programu + další data
   "-XT500_output_filename_69" AT %QB375 : Byte;   // zápid textu v asci pro volbu programu + další data
   "-XT500_output_filename_70" AT %QB376 : Byte;   // zápid textu v asci pro volbu programu + další data
   "-XT500_output_filename_71" AT %QB377 : Byte;   // zápid textu v asci pro volbu programu + další data
   "-XT500_output_filename_72" AT %QB378 : Byte;   // zápid textu v asci pro volbu programu + další data
   "-XT500_output_filename_73" AT %QB379 : Byte;   // zápid textu v asci pro volbu programu + další data
   "-XT500_output_filename_74" AT %QB380 : Byte;   // zápid textu v asci pro volbu programu + další data
   "-XT500_output_filename_75" AT %QB381 : Byte;   // zápid textu v asci pro volbu programu + další data
   "-XT500_output_filename_76" AT %QB382 : Byte;   // zápid textu v asci pro volbu programu + další data
   "-XT500_output_filename_77" AT %QB383 : Byte;   // zápid textu v asci pro volbu programu + další data
   "-XT500_output_filename_78" AT %QB384 : Byte;   // zápid textu v asci pro volbu programu + další data
   "-XT500_output_filename_79" AT %QB385 : Byte;   // zápid textu v asci pro volbu programu + další data
   "-XT500_output_filename_80" AT %QB386 : Byte;   // zápid textu v asci pro volbu programu + další data
   "-XT500_output_filename_81" AT %QB387 : Byte;   // zápid textu v asci pro volbu programu + další data
   "-XT500_output_filename_82" AT %QB388 : Byte;   // zápid textu v asci pro volbu programu + další data
   "-XT500_output_filename_83" AT %QB389 : Byte;   // zápid textu v asci pro volbu programu + další data
   "-XT500_output_filename_84" AT %QB390 : Byte;   // zápid textu v asci pro volbu programu + další data
   "-XT500_output_filename_85" AT %QB391 : Byte;   // zápid textu v asci pro volbu programu + další data
   "-XT500_output_filename_86" AT %QB392 : Byte;   // zápid textu v asci pro volbu programu + další data
   "-XT500_output_filename_87" AT %QB393 : Byte;   // zápid textu v asci pro volbu programu + další data
   "-XT500_output_filename_88" AT %QB394 : Byte;   // zápid textu v asci pro volbu programu + další data
   "-XT500_output_filename_89" AT %QB395 : Byte;   // zápid textu v asci pro volbu programu + další data
   "-XT500_output_filename_90" AT %QB396 : Byte;   // zápid textu v asci pro volbu programu + další data
   "-XT500_output_filename_91" AT %QB397 : Byte;   // zápid textu v asci pro volbu programu + další data
   "-XT500_output_filename_92" AT %QB398 : Byte;   // zápid textu v asci pro volbu programu + další data
   "-XT500_output_filename_93" AT %QB399 : Byte;   // zápid textu v asci pro volbu programu + další data
   "-XT500_output_filename_94" AT %QB400 : Byte;   // zápid textu v asci pro volbu programu + další data
   "-XT500_output_filename_95" AT %QB401 : Byte;   // zápid textu v asci pro volbu programu + další data
   "-XT500_output_filename_96" AT %QB402 : Byte;   // zápid textu v asci pro volbu programu + další data
   "-XT500_output_filename_97" AT %QB403 : Byte;   // zápid textu v asci pro volbu programu + další data
   "-XT500_output_filename_98" AT %QB404 : Byte;   // zápid textu v asci pro volbu programu + další data
   "-XT500_output_filename_99" AT %QB405 : Byte;   // zápid textu v asci pro volbu programu + další data
   "-XT500_output_filename_100" AT %QB406 : Byte;   // zápid textu v asci pro volbu programu + další data
   "-XT500_output_filename_101" AT %QB407 : Byte;   // zápid textu v asci pro volbu programu + další data
   "-XT500_output_filename_102" AT %QB408 : Byte;   // zápid textu v asci pro volbu programu + další data
   "-XT500_output_filename_103" AT %QB409 : Byte;   // zápid textu v asci pro volbu programu + další data
   "-XT500_output_filename_104" AT %QB410 : Byte;   // zápid textu v asci pro volbu programu + další data
   "-XT500_output_filename_105" AT %QB422 : Byte;   // zápid textu v asci pro volbu programu + další data
   "-XT500_output_filename_106" AT %QB423 : Byte;   // zápid textu v asci pro volbu programu + další data
   "-XT500_output_filename_107" AT %QB424 : Byte;   // zápid textu v asci pro volbu programu + další data
   "-XT500_output_filename_108" AT %QB425 : Byte;   // zápid textu v asci pro volbu programu + další data
   "-XT500_output_filename_109" AT %QB426 : Byte;   // zápid textu v asci pro volbu programu + další data
   "-XT500_output_filename_110" AT %QB427 : Byte;   // zápid textu v asci pro volbu programu + další data
   "-XT500_output_filename_111" AT %QB428 : Byte;   // zápid textu v asci pro volbu programu + další data
   "-XT500_output_filename_112" AT %QB429 : Byte;   // zápid textu v asci pro volbu programu + další data
   "-XT500_output_filename_113" AT %QB430 : Byte;   // zápid textu v asci pro volbu programu + další data
   "-XT500_output_filename_114" AT %QB431 : Byte;   // zápid textu v asci pro volbu programu + další data
   "-XT500_output_filename_115" AT %QB432 : Byte;   // zápid textu v asci pro volbu programu + další data
   "-XT500_output_filename_116" AT %QB433 : Byte;   // zápid textu v asci pro volbu programu + další data
   "-XT500_output_filename_117" AT %QB434 : Byte;   // zápid textu v asci pro volbu programu + další data
   "-XT500_output_filename_118" AT %QB435 : Byte;   // zápid textu v asci pro volbu programu + další data
   "-XT500_output_filename_119" AT %QB436 : Byte;   // zápid textu v asci pro volbu programu + další data
   "-XT500_output_filename_120" AT %QB437 : Byte;   // zápid textu v asci pro volbu programu + další data
   "-XT500_output_filename_121" AT %QB438 : Byte;   // zápid textu v asci pro volbu programu + další data
   "-XT500_output_filename_122" AT %QB439 : Byte;   // zápid textu v asci pro volbu programu + další data
   "-XT500_output_filename_123" AT %QB440 : Byte;   // zápid textu v asci pro volbu programu + další data
   "-XT500_output_filename_124" AT %QB441 : Byte;   // zápid textu v asci pro volbu programu + další data
   "-XT500_output_filename_125" AT %QB442 : Byte;   // zápid textu v asci pro volbu programu + další data
   "-XT500_output_filename_126" AT %QB443 : Byte;   // zápid textu v asci pro volbu programu + další data
   "-XT500_output_filename_127" AT %QB444 : Byte;   // zápid textu v asci pro volbu programu + další data
   "-XT500_output_filename_128" AT %QB445 : Byte;   // zápid textu v asci pro volbu programu + další data
   "-XT500_output_filename_129" AT %QB446 : Byte;   // zápid textu v asci pro volbu programu + další data
   "-XT500_output_filename_130" AT %QB447 : Byte;   // zápid textu v asci pro volbu programu + další data
   "-XT500_output_filename_131" AT %QB448 : Byte;   // zápid textu v asci pro volbu programu + další data
   "-XT500_output_filename_132" AT %QB449 : Byte;   // zápid textu v asci pro volbu programu + další data
   "-XT500_output_filename_133" AT %QB450 : Byte;   // zápid textu v asci pro volbu programu + další data
   "-XT500_output_filename_134" AT %QB451 : Byte;   // zápid textu v asci pro volbu programu + další data
   "-XT500_output_filename_135" AT %QB452 : Byte;   // zápid textu v asci pro volbu programu + další data
   "-XT500_output_filename_136" AT %QB453 : Byte;   // zápid textu v asci pro volbu programu + další data
   "-XT500_output_filename_137" AT %QB454 : Byte;   // zápid textu v asci pro volbu programu + další data
   "-XT500_output_filename_138" AT %QB455 : Byte;   // zápid textu v asci pro volbu programu + další data
END_VAR

TYPE "AXIS_FESTO_SIN_POS_TEL_111"
   STRUCT
      AXIS_TEL_111 : Struct
         SENDING : Struct
            MODE_POS : Int;   // JOG = 7 REALATIVE = 2 ABSOLUTNĚ = 1 HOMING = 4 / JOG = 7 RELATIVE = 2 ABSOLUTE = 1 HOMING = 4
            ENABLE_AXIS : Bool;   // ENABLE
            CANCEL_TRAVERSING : Bool;
            INTERMEDIATE_STOP : Bool;
            POSITIVE : Bool;
            NEGATIVE : Bool;
            JOG_1 : Bool;
            JOG_2 : Bool;
            FLI_REF : Bool;
            ACK_ERROR : Bool;
            EXECUTE_MODE : Bool;
            POSITION : DInt;
            VELOCITY : DInt;
            OVER_V : Int;
            OVER_ACC : Int;
            OVER_DEC : Int;
         END_STRUCT;
         READ : Struct
            AXIS_ENABLED : Bool;
            AXIS_POS_OK : Bool;
            AXIS_SP_FIXED : Bool;
            AXIS_REF : Bool;
            AXIS_WARN : Bool;
            AXIS_ERROR : Bool;
            LOCKOUT : Bool;
            ACT_VELOCITY : DInt;
            ACT_POSITION : DInt;
            ACT_MODE : Int;
            EPOS_ZSW_1 : Word;
            EPOS_ZSW_2 : Word;
            ACT_WARN : Word;
            ACT_FAULT : Word;
            ERROR : Bool;
            STATUS : Word;
            DIAGLD : Word;
         END_STRUCT;
      END_STRUCT;
   END_STRUCT;
END_TYPE

TYPE "AXIS_VIRT_N_CODE"
   STRUCT
      AXIS : Struct
         SENDING : Struct
            MC_POWER { ExternalAccessible := 'False'; ExternalVisible := 'False'; ExternalWritable := 'False'} : Struct
               ENABLE : Bool;
               START_MODE : Int;
               STOP_MODE : Int;
            END_STRUCT;
            MC_HOME { ExternalAccessible := 'False'; ExternalVisible := 'False'; ExternalWritable := 'False'} : Struct
               EXECUTE : Bool;
               POSITION : Real;
               MODE : Int;
            END_STRUCT;
            MC_MOVE_JOG { ExternalAccessible := 'False'; ExternalVisible := 'False'; ExternalWritable := 'False'} : Struct
               JOG_FORWARD : Bool;
               JOG_BACKWARD : Bool;
               VELOCITY : Real;
               POSITION_CONTROLED : Bool;
            END_STRUCT;
            MC_RESET { ExternalAccessible := 'False'; ExternalVisible := 'False'; ExternalWritable := 'False'} : Struct
               EXECUTE : Bool;
               RESTART : Bool;
            END_STRUCT;
            MC_MOVE_ABSOLUTE_JOG { ExternalAccessible := 'False'; ExternalVisible := 'False'; ExternalWritable := 'False'} : Struct
               EXECUTE : Bool;
               POSITION : Real;
               VELOCITY : Real;
               DIRECTION : Int;
            END_STRUCT;
            MC_HALT { ExternalAccessible := 'False'; ExternalVisible := 'False'; ExternalWritable := 'False'} : Struct
               EXECUTE : Bool;
            END_STRUCT;
         END_STRUCT;
         READ : Struct
            MC_POWER : Struct
               STATUS : Bool;
               BUSY : Bool;
               ERROR : Bool;
               ERROR_ID : Word;
               ERROR_INTO : Word;
            END_STRUCT;
            MC_HOME : Struct
               DONE : Bool;
               BUSY : Bool;
               COMAND_ABORTED : Bool;
               ERROR : Bool;
               ERROR_ID : Word;
               ERROR_INTO : Word;
               REFERENCE_MARK_POSITION : Real;
            END_STRUCT;
            MC_MOVE_JOG : Struct
               IN_VELOCITY : Bool;
               BUSY : Bool;
               COMAND_ABORTED : Bool;
               ERROR : Bool;
               ERROR_ID : Word;
               ERROR_INTO : Word;
            END_STRUCT;
            MC_RESET : Struct
               DONE : Bool;
               BUSY : Bool;
               ERROR : Bool;
               ERROR_ID : Word;
               ERROR_INTO : Word;
            END_STRUCT;
            MC_MOVE_ABSOLUTE : Struct
               DONE : Bool;
               BYSY : Bool;
               COMAND_ABORTED : Bool;
               ERROR : Bool;
               ERROR_ID : Word;
               ERROR_INTO : Word;
            END_STRUCT;
            MC_HALT : Struct
               done : Bool;
               BUSY : Bool;
               error : Bool;
               COMAD_ABORTED : Bool;
               ERROR_ID : Word;
               ERROR_INTO : Word;
            END_STRUCT;
         END_STRUCT;
      END_STRUCT;
   END_STRUCT;
END_TYPE

TYPE "DATA_RECEPT"
   STRUCT
      NUMBER_PROG { S7_SetPoint := 'True'} : Int;
      PROG_NAME { S7_SetPoint := 'True'} : String[38];
      OS_Z { S7_SetPoint := 'True'} : DInt;
      SELECTED : Bool;
   END_STRUCT;
END_TYPE

TYPE "TDiag_StatusExt"
   STRUCT
      Interfaceld : HW_ANY;
      ID : CONN_OUC;
      ConnectionType : Byte;
      ActivateEstablished : Bool;
      State : Byte;
      Kind : Byte;
      SentBytes : UDInt;
      ReceivedBytes : UDInt;
   END_STRUCT;
END_TYPE

TYPE "T_CON_DATA"
   STRUCT
      TCON : Struct
         IN : Struct
            START : Bool;
            ID : CONN_OUC;
         END_STRUCT;
         OUT : Struct
            DONE : Bool;
            BYSY : Bool;
            ERROR : Bool;
            STATUS : Word;
         END_STRUCT;
      END_STRUCT;
   END_STRUCT;
END_TYPE

TYPE "T_DISCON_DATA"
   STRUCT
      TDISCON : Struct
         IN : Struct
            DISCONNECT : Bool;
            ID : CONN_OUC;
         END_STRUCT;
         OUT : Struct
            DONE : Bool;
            BUSY : Bool;
            ERROR : Bool;
            STATUS : Word;
         END_STRUCT;
      END_STRUCT;
   END_STRUCT;
END_TYPE

TYPE "T_RCV_DATA"
   STRUCT
      TRCV : Struct
         IN : Struct
            READ : Bool;
            ID : CONN_OUC;
            LEN : UDInt;
            ADHOC : Bool;
            DATA : Array[0..254] of Char;
         END_STRUCT;
         OUT : Struct
            NDR : Bool;
            BYSY : Bool;
            ERROR : Bool;
            STATUS : Word;
            RCVD_LEN : DWord;
         END_STRUCT;
      END_STRUCT;
   END_STRUCT;
END_TYPE

DATA_BLOCK "DB_HMI_recype"   // DB2
{ S7_Optimized_Access := 'TRUE' }
// stored: MemoryReserve 100
   VAR
      recipe : Struct
         Zprava : Int := 2;   // dvoumístné číslo přeneseno a doplněno po bytech do šablony zprávy
         PRG_CAM_etiketa : Int := 1;   // program v kameře která kontroluje papír co se vkládá pod folii
         PRG_CAM_folie : Int;   // kamery kontrolující folii
         vyrazovac_on_off : Bool := true;   // false - neposílat signál pro vyřazovač
         variabilni_pole_on_off : Bool := true;   // false - neposílat variabilní pole
         pole_string_1 : String[20] := 'Ceska republika';   // textove_pole - není bráno z receptůry ale volně zadatalné
         pole_string_2 : String[10];   // textove_pole - není bráno z receptůry ale volně zadatalné
      END_STRUCT;
      fronta : Array[1..5] of Struct
         prenaseny_text : String[100];   // načtený text kamerou
         balik_den : Int;   // aktualni číslo plata
         vyrazeni : Bool;   // vyřazení
      END_STRUCT;
      obsazenost_fronty : Int;
      ODESLI_dATA : Bool;
      VZDALENOST_KAMERA_ETIKETA_POZADOVANA : DInt := 20;
      VZDALENOST_KAMERY_FOLIE_POZADOVANA : DInt := 150;
      meze : DInt := 35;
      aktualni_poloha : DInt;
   END_VAR
BEGIN
END_DATA_BLOCK

DATA_BLOCK "DB_data_ctena"   // DB7
{ S7_Optimized_Access := 'TRUE' }
// stored: MemoryReserve 100
   VAR
      array_of_byte : Array[0..150] of Byte;
      array_of_char : Array[0..150] of Char;
      cteny_string : String[150];
      upraveny : String[150];
   END_VAR
BEGIN
END_DATA_BLOCK

DATA_BLOCK "DB_prikazy_tiskarna"   // DB4
{ S7_Optimized_Access := 'TRUE' }
// stored: MemoryReserve 0
   VAR
      task : Array[0..6, 0..255] of Byte;
      DATA : Array[0..255] of Byte;
      ADRESACE_POLE : Int := 1;
      hodnota_pamet : Int := 1;
      cislo_zpravy : Int := 2;   // zpráva má pevný formát mění se pouze číslo které je odesíláno jako string před převedením do stringu je rozseknuto na byte a kopírováno jako jednotlyvý znak
      DATA_RECIVR : Array[0..255] of Byte;
      byte_1 : Byte := 16#30;
      byte_2 : Byte := 16#32;
      text_pole_1 : String[30];   // pole jedno - odkud pochází
      text_pole_2 : String[10];   // pole dvě - datum spotřeby požadovaný formát xx.xx.xxxx
   END_VAR
BEGIN
   task[0,0] := 16#00;   // get_status
   task[0,1..4] := 16#00;
   task[0,5] := 16#06;
   task[0,6] := 16#01;
   task[0,7] := 16#64;
   task[0,8] := 16#00;
   task[0,9] := 16#02;
   task[0,10] := 16#01;
   task[0,11] := 16#45;
   // task[0,255] : get_status
   task[1,0] := 16#00;   // START_TISKU
   task[1,1] := 16#00;   // START_TISKU
   task[1,2] := 16#00;   // START_TISKU
   task[1,3] := 16#00;   // START_TISKU
   task[1,4] := 16#00;   // START_TISKU
   task[1,5] := 16#0D;   // START_TISKU
   task[1,6] := 16#01;   // START_TISKU
   task[1,7] := 16#64;   // START_TISKU
   task[1,8] := 16#00;   // START_TISKU
   task[1,9] := 16#09;   // START_TISKU
   task[1,10] := 16#01;   // START_TISKU
   task[1,11] := 16#20;   // START_TISKU
   task[1,12] := 16#02;   // START_TISKU
   task[1,13] := 16#13;   // START_TISKU
   task[1,14] := 16#00;   // START_TISKU
   task[1,15] := 16#00;   // START_TISKU
   task[1,16] := 16#00;   // START_TISKU
   task[1,17] := 16#00;   // START_TISKU
   task[1,18] := 16#00;   // START_TISKU
   // task[1,255] : START_TISKU
   task[2,0] := 16#00;   // STOP_TISKU
   task[2,1] := 16#00;   // STOP_TISKU
   task[2,2] := 16#00;   // STOP_TISKU
   task[2,3] := 16#00;   // STOP_TISKU
   task[2,4] := 16#00;   // STOP_TISKU
   task[2,5] := 16#0D;   // STOP_TISKU
   task[2,6] := 16#01;   // STOP_TISKU
   task[2,7] := 16#64;   // STOP_TISKU
   task[2,8] := 16#00;   // STOP_TISKU
   task[2,9] := 16#09;   // STOP_TISKU
   task[2,10] := 16#01;   // STOP_TISKU
   task[2,11] := 16#20;   // STOP_TISKU
   task[2,12] := 16#02;   // STOP_TISKU
   task[2,13] := 16#13;   // STOP_TISKU
   task[2,14] := 16#00;   // STOP_TISKU
   task[2,15] := 16#00;   // STOP_TISKU
   task[2,16] := 16#00;   // STOP_TISKU
   task[2,17] := 16#00;   // STOP_TISKU
   task[2,18] := 16#01;   // STOP_TISKU
   // task[2,19] : STOP_TISKU
   // task[2,20] : STOP_TISKU
   // task[2,21] : STOP_TISKU
   task[3,0] := 16#00;
   task[3,1] := 16#00;   // VÝBĚR ZPRÁVY
   task[3,2] := 16#00;   // VÝBĚR ZPRÁVY
   task[3,3] := 16#00;   // VÝBĚR ZPRÁVY
   task[3,4] := 16#00;
   task[3,5] := 16#1A;
   task[3,6] := 16#01;
   task[3,7] := 16#64;
   task[3,8] := 16#00;
   task[3,9] := 16#16;
   task[3,10] := 16#01;
   task[3,11] := 16#20;
   task[3,12] := 16#02;
   task[3,13] := 16#4C;
   task[3,14..18] := 16#00;
   task[3,19] := 16#0C;
   task[3,20] := 16#4D;
   task[3,21] := 16#53;
   task[3,22] := 16#47;
   task[3,23..25] := 16#30;
   task[3,28] := 16#2E;
   task[3,29] := 16#78;
   task[3,30] := 16#6D;
   task[3,31] := 16#6C;
   task[4,0] := 16#00;   // VYPLNĚNÍ DAT MAX 30 ZNAKŮ DO JEDNOHO POLE AKTUÁLNĚ
   task[4,1] := 16#00;   // VYPLNĚNÍ DAT MAX 30 ZNAKŮ DO JEDNOHO POLE AKTUÁLNĚ
   task[4,2] := 16#00;   // VYPLNĚNÍ DAT MAX 30 ZNAKŮ DO JEDNOHO POLE AKTUÁLNĚ
   task[4,3] := 16#00;   // VYPLNĚNÍ DAT MAX 30 ZNAKŮ DO JEDNOHO POLE AKTUÁLNĚ
   task[4,4] := 16#00;   // VYPLNĚNÍ DAT MAX 30 ZNAKŮ DO JEDNOHO POLE AKTUÁLNĚ
   task[4,5] := 16#3C;   // VYPLNĚNÍ DAT MAX 30 ZNAKŮ DO JEDNOHO POLE AKTUÁLNĚ
   task[4,6] := 16#01;   // VYPLNĚNÍ DAT MAX 30 ZNAKŮ DO JEDNOHO POLE AKTUÁLNĚ
   task[4,7] := 16#64;   // VYPLNĚNÍ DAT MAX 30 ZNAKŮ DO JEDNOHO POLE AKTUÁLNĚ
   task[4,8] := 16#00;   // VYPLNĚNÍ DAT MAX 30 ZNAKŮ DO JEDNOHO POLE AKTUÁLNĚ
   task[4,9] := 16#38;   // VYPLNĚNÍ DAT MAX 30 ZNAKŮ DO JEDNOHO POLE AKTUÁLNĚ
   task[4,10] := 16#01;   // VYPLNĚNÍ DAT MAX 30 ZNAKŮ DO JEDNOHO POLE AKTUÁLNĚ
   task[4,11] := 16#CF;   // VYPLNĚNÍ DAT MAX 30 ZNAKŮ DO JEDNOHO POLE AKTUÁLNĚ
   task[4,12] := 16#00;   // VYPLNĚNÍ DAT MAX 30 ZNAKŮ DO JEDNOHO POLE AKTUÁLNĚ
   task[4,13] := 16#00;   // VYPLNĚNÍ DAT MAX 30 ZNAKŮ DO JEDNOHO POLE AKTUÁLNĚ
   task[4,14] := 16#00;   // VYPLNĚNÍ DAT MAX 30 ZNAKŮ DO JEDNOHO POLE AKTUÁLNĚ
   task[4,15] := 16#00;
   task[4,16] := 16#1E;
   task[4,17] := 16#51;
   task[4,18] := 16#57;
   task[4,19] := 16#45;
   task[4,20] := 16#52;
   task[4,21] := 16#54;
   task[4,22] := 16#5A;
   task[4,23] := 16#55;
   task[4,24] := 16#49;
   task[4,25] := 16#4F;
   task[4,26] := 16#50;
   task[4,27] := 16#41;
   task[4,28] := 16#53;
   task[4,29] := 16#44;
   task[4,30] := 16#46;
   task[4,31] := 16#47;
   task[4,32] := 16#48;
   task[4,33] := 16#4A;
   task[4,34] := 16#4B;
   task[4,35] := 16#4C;
   task[4,36] := 16#59;
   task[4,37] := 16#58;
   task[4,38] := 16#43;
   task[4,39] := 16#56;
   task[4,40] := 16#42;
   task[4,41] := 16#4E;
   task[4,42] := 16#4D;
   task[4,43] := 16#31;
   task[4,44] := 16#32;
   task[4,45] := 16#33;
   task[4,46] := 16#34;
   task[4,47..65] := 16#00;
   task[6,0] := 16#00;   // SMAZANÍ A PŘENASTAVENÍ ABY TISKÁRNA NEBAFROVALA ALE TISKLA ODESLANÁ DATA DO KOLA
   task[6,1] := 16#00;   // SMAZANÍ A PŘENASTAVENÍ ABY TISKÁRNA NEBAFROVALA ALE TISKLA ODESLANÁ DATA DO KOLA
   task[6,2] := 16#00;   // SMAZANÍ A PŘENASTAVENÍ ABY TISKÁRNA NEBAFROVALA ALE TISKLA ODESLANÁ DATA DO KOLA
   task[6,3] := 16#00;   // SMAZANÍ A PŘENASTAVENÍ ABY TISKÁRNA NEBAFROVALA ALE TISKLA ODESLANÁ DATA DO KOLA
   task[6,4] := 16#00;   // SMAZANÍ A PŘENASTAVENÍ ABY TISKÁRNA NEBAFROVALA ALE TISKLA ODESLANÁ DATA DO KOLA
   task[6,5] := 16#0D;   // SMAZANÍ A PŘENASTAVENÍ ABY TISKÁRNA NEBAFROVALA ALE TISKLA ODESLANÁ DATA DO KOLA
   task[6,6] := 16#01;   // SMAZANÍ A PŘENASTAVENÍ ABY TISKÁRNA NEBAFROVALA ALE TISKLA ODESLANÁ DATA DO KOLA
   task[6,7] := 16#64;   // SMAZANÍ A PŘENASTAVENÍ ABY TISKÁRNA NEBAFROVALA ALE TISKLA ODESLANÁ DATA DO KOLA
   task[6,8] := 16#00;
   task[6,9] := 16#09;
   task[6,10] := 16#01;
   task[6,11] := 16#CE;
   task[6,12..17] := 16#00;
   task[6,18] := 16#01;
   // DATA_RECIVR[0] : 16#00
   // DATA_RECIVR[1] : 16#00
   // DATA_RECIVR[2] : 16#00
   // DATA_RECIVR[3] : 16#00
   // DATA_RECIVR[4] : 16#00
   // DATA_RECIVR[5] : 16#06
   // DATA_RECIVR[6] : 16#01
   // DATA_RECIVR[7] : 16#64
   // DATA_RECIVR[8] : 16#00
   // DATA_RECIVR[9] : 16#02
   // DATA_RECIVR[10] : 16#01
   // DATA_RECIVR[11] : 16#4F
   // DATA_RECIVR[12] : 16#00
   // DATA_RECIVR[13] : 16#00
   // DATA_RECIVR[14] : 16#00
   // DATA_RECIVR[15] : 16#00
   // DATA_RECIVR[16] : 16#00
   // DATA_RECIVR[17] : 16#06
   // DATA_RECIVR[18] : 16#01
   // DATA_RECIVR[19] : 16#64
   // DATA_RECIVR[20] : 16#00
   // DATA_RECIVR[21] : 16#02
   // DATA_RECIVR[22] : 16#01
   // DATA_RECIVR[23] : 16#4F
   // DATA_RECIVR[24] : 16#00
   // DATA_RECIVR[25] : 16#00
   // DATA_RECIVR[26] : 16#00
   // DATA_RECIVR[27] : 16#00
   // DATA_RECIVR[28] : 16#00
   // DATA_RECIVR[29] : 16#06
   // DATA_RECIVR[30] : 16#01
   // DATA_RECIVR[31] : 16#64
   // DATA_RECIVR[32] : 16#00
   // DATA_RECIVR[33] : 16#02
   // DATA_RECIVR[34] : 16#01
   // DATA_RECIVR[35] : 16#4F
   // DATA_RECIVR[36] : 16#00
   // DATA_RECIVR[37] : 16#00
   // DATA_RECIVR[38] : 16#00
   // DATA_RECIVR[39] : 16#00
   // DATA_RECIVR[40] : 16#00
   // DATA_RECIVR[41] : 16#06
   // DATA_RECIVR[42] : 16#01
   // DATA_RECIVR[43] : 16#64
   // DATA_RECIVR[44] : 16#00
   // DATA_RECIVR[45] : 16#02
   // DATA_RECIVR[46] : 16#01
   // DATA_RECIVR[47] : 16#4F
   // DATA_RECIVR[48] : 16#00
   // DATA_RECIVR[49] : 16#00
   // DATA_RECIVR[50] : 16#00
   // DATA_RECIVR[51] : 16#00
   // DATA_RECIVR[52] : 16#00
   // DATA_RECIVR[53] : 16#06
   // DATA_RECIVR[54] : 16#01
   // DATA_RECIVR[55] : 16#64
   // DATA_RECIVR[56] : 16#00
   // DATA_RECIVR[57] : 16#02
   // DATA_RECIVR[58] : 16#01
   // DATA_RECIVR[59] : 16#4F
   // DATA_RECIVR[60] : 16#00
   // DATA_RECIVR[61] : 16#00
   // DATA_RECIVR[62] : 16#00
   // DATA_RECIVR[63] : 16#00
   // DATA_RECIVR[64] : 16#00
   // DATA_RECIVR[65] : 16#06
   // DATA_RECIVR[66] : 16#01
   // DATA_RECIVR[67] : 16#64
   // DATA_RECIVR[68] : 16#00
   // DATA_RECIVR[69] : 16#02
   // DATA_RECIVR[70] : 16#01
   // DATA_RECIVR[71] : 16#4F
   // DATA_RECIVR[72] : 16#00
   // DATA_RECIVR[73] : 16#00
   // DATA_RECIVR[74] : 16#00
   // DATA_RECIVR[75] : 16#00
   // DATA_RECIVR[76] : 16#00
   // DATA_RECIVR[77] : 16#06
   // DATA_RECIVR[78] : 16#01
   // DATA_RECIVR[79] : 16#64
   // DATA_RECIVR[80] : 16#00
   // DATA_RECIVR[81] : 16#02
   // DATA_RECIVR[82] : 16#01
   // DATA_RECIVR[83] : 16#4F
   // DATA_RECIVR[84] : 16#00
   // DATA_RECIVR[85] : 16#00
   // DATA_RECIVR[86] : 16#00
   // DATA_RECIVR[87] : 16#00
   // DATA_RECIVR[88] : 16#00
   // DATA_RECIVR[89] : 16#06
   // DATA_RECIVR[90] : 16#01
   // DATA_RECIVR[91] : 16#64
   // DATA_RECIVR[92] : 16#00
   // DATA_RECIVR[93] : 16#02
   // DATA_RECIVR[94] : 16#01
   // DATA_RECIVR[95] : 16#4F
   // DATA_RECIVR[96] : 16#00
   // DATA_RECIVR[97] : 16#00
   // DATA_RECIVR[98] : 16#00
   // DATA_RECIVR[99] : 16#00
   // DATA_RECIVR[100] : 16#00
   // DATA_RECIVR[101] : 16#06
   // DATA_RECIVR[102] : 16#01
   // DATA_RECIVR[103] : 16#64
   // DATA_RECIVR[104] : 16#00
   // DATA_RECIVR[105] : 16#02
   // DATA_RECIVR[106] : 16#01
   // DATA_RECIVR[107] : 16#4F
   // DATA_RECIVR[108] : 16#00
   // DATA_RECIVR[109] : 16#00
   // DATA_RECIVR[110] : 16#00
   // DATA_RECIVR[111] : 16#00
   // DATA_RECIVR[112] : 16#00
   // DATA_RECIVR[113] : 16#06
   // DATA_RECIVR[114] : 16#01
   // DATA_RECIVR[115] : 16#64
   // DATA_RECIVR[116] : 16#00
   // DATA_RECIVR[117] : 16#02
   // DATA_RECIVR[118] : 16#01
   // DATA_RECIVR[119] : 16#4F
   // DATA_RECIVR[120] : 16#00
   // DATA_RECIVR[121] : 16#00
   // DATA_RECIVR[122] : 16#00
   // DATA_RECIVR[123] : 16#00
   // DATA_RECIVR[124] : 16#00
   // DATA_RECIVR[125] : 16#06
   // DATA_RECIVR[126] : 16#01
   // DATA_RECIVR[127] : 16#64
   // DATA_RECIVR[128] : 16#00
   // DATA_RECIVR[129] : 16#02
   // DATA_RECIVR[130] : 16#01
   // DATA_RECIVR[131] : 16#4F
   // DATA_RECIVR[132] : 16#00
   // DATA_RECIVR[133] : 16#00
   // DATA_RECIVR[134] : 16#00
   // DATA_RECIVR[135] : 16#00
   // DATA_RECIVR[136] : 16#00
   // DATA_RECIVR[137] : 16#06
   // DATA_RECIVR[138] : 16#01
   // DATA_RECIVR[139] : 16#64
   // DATA_RECIVR[140] : 16#00
   // DATA_RECIVR[141] : 16#02
   // DATA_RECIVR[142] : 16#01
   // DATA_RECIVR[143] : 16#4F
   // DATA_RECIVR[144] : 16#00
   // DATA_RECIVR[145] : 16#00
   // DATA_RECIVR[146] : 16#00
   // DATA_RECIVR[147] : 16#00
   // DATA_RECIVR[148] : 16#00
   // DATA_RECIVR[149] : 16#06
   // DATA_RECIVR[150] : 16#01
   // DATA_RECIVR[151] : 16#64
   // DATA_RECIVR[152] : 16#00
   // DATA_RECIVR[153] : 16#02
   // DATA_RECIVR[154] : 16#01
   // DATA_RECIVR[155] : 16#4F
   // DATA_RECIVR[156] : 16#00
   // DATA_RECIVR[157] : 16#00
   // DATA_RECIVR[158] : 16#00
   // DATA_RECIVR[159] : 16#00
   // DATA_RECIVR[160] : 16#00
   // DATA_RECIVR[161] : 16#06
   // DATA_RECIVR[162] : 16#01
   // DATA_RECIVR[163] : 16#64
   // DATA_RECIVR[164] : 16#00
   // DATA_RECIVR[165] : 16#02
   // DATA_RECIVR[166] : 16#01
   // DATA_RECIVR[167] : 16#4F
   // DATA_RECIVR[168] : 16#00
   // DATA_RECIVR[169] : 16#00
   // DATA_RECIVR[170] : 16#00
   // DATA_RECIVR[171] : 16#00
   // DATA_RECIVR[172] : 16#00
   // DATA_RECIVR[173] : 16#06
   // DATA_RECIVR[174] : 16#01
   // DATA_RECIVR[175] : 16#64
   // DATA_RECIVR[176] : 16#00
   // DATA_RECIVR[177] : 16#02
   // DATA_RECIVR[178] : 16#01
   // DATA_RECIVR[179] : 16#4F
   // DATA_RECIVR[180] : 16#00
   // DATA_RECIVR[181] : 16#00
   // DATA_RECIVR[182] : 16#00
   // DATA_RECIVR[183] : 16#00
   // DATA_RECIVR[184] : 16#00
   // DATA_RECIVR[185] : 16#06
   // DATA_RECIVR[186] : 16#01
   // DATA_RECIVR[187] : 16#64
   // DATA_RECIVR[188] : 16#00
   // DATA_RECIVR[189] : 16#02
   // DATA_RECIVR[190] : 16#01
   // DATA_RECIVR[191] : 16#4F
   // DATA_RECIVR[192] : 16#00
   // DATA_RECIVR[193] : 16#00
   // DATA_RECIVR[194] : 16#00
   // DATA_RECIVR[195] : 16#00
   // DATA_RECIVR[196] : 16#00
   // DATA_RECIVR[197] : 16#06
   // DATA_RECIVR[198] : 16#01
   // DATA_RECIVR[199] : 16#64
   // DATA_RECIVR[200] : 16#00
   // DATA_RECIVR[201] : 16#02
   // DATA_RECIVR[202] : 16#01
   // DATA_RECIVR[203] : 16#4F
   // DATA_RECIVR[204] : 16#00
   // DATA_RECIVR[205] : 16#00
   // DATA_RECIVR[206] : 16#00
   // DATA_RECIVR[207] : 16#00
   // DATA_RECIVR[208] : 16#00
   // DATA_RECIVR[209] : 16#06
   // DATA_RECIVR[210] : 16#01
   // DATA_RECIVR[211] : 16#64
   // DATA_RECIVR[212] : 16#00
   // DATA_RECIVR[213] : 16#02
   // DATA_RECIVR[214] : 16#01
   // DATA_RECIVR[215] : 16#4F
   // DATA_RECIVR[216] : 16#00
   // DATA_RECIVR[217] : 16#00
   // DATA_RECIVR[218] : 16#00
   // DATA_RECIVR[219] : 16#00
   // DATA_RECIVR[220] : 16#00
   // DATA_RECIVR[221] : 16#06
   // DATA_RECIVR[222] : 16#01
   // DATA_RECIVR[223] : 16#64
   // DATA_RECIVR[224] : 16#00
   // DATA_RECIVR[225] : 16#02
   // DATA_RECIVR[226] : 16#01
   // DATA_RECIVR[227] : 16#4F
   // DATA_RECIVR[228] : 16#00
   // DATA_RECIVR[229] : 16#00
   // DATA_RECIVR[230] : 16#00
   // DATA_RECIVR[231] : 16#00
   // DATA_RECIVR[232] : 16#00
   // DATA_RECIVR[233] : 16#07
   // DATA_RECIVR[234] : 16#01
   // DATA_RECIVR[235] : 16#64
   // DATA_RECIVR[236] : 16#00
   // DATA_RECIVR[237] : 16#03
   // DATA_RECIVR[238] : 16#01
   // DATA_RECIVR[239] : 16#31
   // DATA_RECIVR[240] : 16#04
   // DATA_RECIVR[241] : 16#00
   // DATA_RECIVR[242] : 16#00
   // DATA_RECIVR[243] : 16#00
   // DATA_RECIVR[244] : 16#00
   // DATA_RECIVR[245] : 16#00
   // DATA_RECIVR[246] : 16#07
   // DATA_RECIVR[247] : 16#01
   // DATA_RECIVR[248] : 16#64
   // DATA_RECIVR[249] : 16#00
   // DATA_RECIVR[250] : 16#03
   // DATA_RECIVR[251] : 16#01
   // DATA_RECIVR[252] : 16#45
   // DATA_RECIVR[253] : 16#00
   // DATA_RECIVR[254] : 16#00
   // DATA_RECIVR[255] : 16#00
END_DATA_BLOCK

DATA_BLOCK "DB_SYSTEM"   // DB12
{ S7_Optimized_Access := 'TRUE' }
// stored: MemoryReserve 100
   VAR RETAIN
      OP2 : Struct
         M1 { S7_SetPoint := 'True'} : Time;
         M2 { S7_SetPoint := 'True'} : Time;
         M3 { S7_SetPoint := 'True'} : Time;
         M4 { S7_SetPoint := 'True'} : Time;
         M5 { S7_SetPoint := 'True'} : Time;
         M6 { S7_SetPoint := 'True'} : Time;
         M7 { S7_SetPoint := 'True'} : Time;
         M8 { S7_SetPoint := 'True'} : Time;
      END_STRUCT;
      OP3 : Struct
         M1 { S7_SetPoint := 'True'} : Time;
         M2 { S7_SetPoint := 'True'} : Time;
         M3 { S7_SetPoint := 'True'} : Time;
         M4 { S7_SetPoint := 'True'} : Time;
         M5 { S7_SetPoint := 'True'} : Time;
         M6 { S7_SetPoint := 'True'} : Time;
         M7 { S7_SetPoint := 'True'} : Time;
         M8 { S7_SetPoint := 'True'} : Time;
      END_STRUCT;
   END_VAR
BEGIN
END_DATA_BLOCK

DATA_BLOCK "DB_Manual"   // DB8
{ S7_Optimized_Access := 'TRUE' }
// stored: MemoryReserve 100
   VAR
      xManEtiketa : Bool;   // TRUE = světla + trigger etiketa
      xManFolie : Bool;   // TRUE = světla + trigger folie
      test_vyr : Bool;
   END_VAR
BEGIN
END_DATA_BLOCK

